(* IEC 61131-3 sources: plc-st-coding-agent/progress/evidence/f14_v11_public_20261113/jobs/custom_deepseek-v4pro (part 3) *)

(* ---- public-hard-04.raw_candidate_04.st ---- *)
(* ENGINEERING_CONTRACT
   elementCount DINT: retained process value; 0 after reset, +1 successful enqueue, -1 successful dequeue, held otherwise; range 0..capacity.
   status WORD: overwritten every invocation; 0 idle/reset/success, 16#8002 rejected full enqueue, 16#8001 rejected empty dequeue; reset priority sets 0.
   queue state: first invocation empty; reset priority clears head/tail/count; enqueue writes at tail, dequeue reads head; indices 0..capacity-1.
   edge triggers: R_TRIG consumed every scan; reset priority ignores edge requests; simultaneous enqueue+dequeue unspecified -> no-op.
   units/boundaries: capacity positive DINT derived once from buffer size / item element size; element copied byte-wise from item address.
*)
(* CONTRACT_RULES [] *)
FUNCTION_BLOCK FIFO
VAR_INPUT
    enqueue : BOOL;
    dequeue : BOOL;
    reset : BOOL;
END_VAR
VAR_OUTPUT
    elementCount : DINT;
    status : WORD;
END_VAR
VAR_IN_OUT
    item : VARIANT;
    buffer : VARIANT;
END_VAR
VAR
    local_rEnq : R_TRIG;
    local_rDeq : R_TRIG;
    local_enqEdge : BOOL;
    local_deqEdge : BOOL;

    local_associated : BOOL := FALSE;
    local_pBufferBase : POINTER TO BYTE;
    local_pItemBase : POINTER TO BYTE;
    local_elemSize : DINT := 1;
    local_capacity : DINT := 1;

    local_count : DINT := 0;
    local_head : DINT := 0;
    local_tail : DINT := 0;

    local_bufInfo : __SYSTEM.VAR_INFO;
    local_itemInfo : __SYSTEM.VAR_INFO;

    local_pSrc : POINTER TO BYTE;
    local_pDst : POINTER TO BYTE;
    local_offset : DINT;
    local_copiedBytes : UDINT;
END_VAR

(* Consume rising edges every scan so reset cannot create ghost operations later. *)
local_rEnq(CLK := enqueue);
local_enqEdge := local_rEnq.Q;
local_rDeq(CLK := dequeue);
local_deqEdge := local_rDeq.Q;

status := 16#0000;

(* One-time association of buffer and item storage, using the first invocation. *)
IF NOT local_associated THEN
    local_bufInfo := __VARINFO(buffer);
    local_itemInfo := __VARINFO(item);

    local_elemSize := local_itemInfo.diSize;
    IF local_elemSize <= 0 THEN
        local_elemSize := 1;
    END_IF;

    local_capacity := local_bufInfo.diSize / local_elemSize;
    IF local_capacity < 1 THEN
        local_capacity := 1;
    END_IF;

    local_pBufferBase := local_bufInfo.pvAddress;
    local_pItemBase := local_itemInfo.pvAddress;
    local_associated := TRUE;
END_IF;

IF reset THEN
    (* Reset has priority over all operations; stored values remain untouched. *)
    local_count := 0;
    local_head := 0;
    local_tail := 0;
    status := 16#0000;
ELSE
    IF local_enqEdge AND NOT local_deqEdge THEN
        IF local_count < local_capacity THEN
            (* Copy current item value into tail slot. *)
            local_pSrc := local_pItemBase;
            local_pDst := local_pBufferBase;
            local_offset := local_tail * local_elemSize;
            local_pDst := local_pDst + local_offset;
            local_copiedBytes := SysMemCpy(
                pbyDest := local_pDst,
                pbySource := local_pSrc,
                dwCount := TO_DWORD(local_elemSize)
            );

            local_tail := (local_tail + 1) MOD local_capacity;
            local_count := local_count + 1;
            status := 16#0000;
        ELSE
            status := 16#8002; (* enqueue rejected: full *)
        END_IF;
    ELSIF local_deqEdge AND NOT local_enqEdge THEN
        IF local_count > 0 THEN
            (* Copy head element back to item. *)
            local_pSrc := local_pBufferBase;
            local_offset := local_head * local_elemSize;
            local_pSrc := local_pSrc + local_offset;
            local_pDst := local_pItemBase;
            local_copiedBytes := SysMemCpy(
                pbyDest := local_pDst,
                pbySource := local_pSrc,
                dwCount := TO_DWORD(local_elemSize)
            );

            local_head := (local_head + 1) MOD local_capacity;
            local_count := local_count - 1;
            status := 16#0000;
        ELSE
            status := 16#8001; (* dequeue rejected: empty *)
        END_IF;
    END_IF;
END_IF;

elementCount := local_count;
END_FUNCTION_BLOCK

(* ---- public-hard-05.candidate_01.st ---- *)
(* ENGINEERING_CONTRACT
Manual: moving/grip/release outputs are combinational from corresponding button AND NOT corresponding limit switch; releasing the button clears the output. PUB001, PUB005.
SingleStep: rising Start advances only when idle or current step limit reached; each step holds its output until its limit, then waits for next Start. After step 8, next Start goes to step 1. PUB002.
SingleCycle: rising Start starts step 1; each step auto-advances on its completion limit, then stops at step 0 after step 8. PUB003.
Continuous: rising Start starts step 1; auto-advances and loops 8->1. PUB004.
EmergencyStop=FALSE forces all outputs FALSE and freezes automatic state changes. No reset is inferred. PUB005.
Completion feedback uses DownLimitSwitch, UpLimitSwitch, LeftLimitSwitch, RightLimitSwitch, GripLimitSwitch, ReleaseLimitSwitch. Unspecified mode-change behavior preserves the automatic step state.
*)
(* CONTRACT_RULES [] *)
FUNCTION_BLOCK FB_MechanicalArmControl
VAR CONSTANT
    cStepDown1 : INT := 1;
    cStepGrip : INT := 2;
    cStepUp1 : INT := 3;
    cStepRight : INT := 4;
    cStepDown2 : INT := 5;
    cStepRelease : INT := 6;
    cStepUp2 : INT := 7;
    cStepLeft : INT := 8;
END_VAR
VAR
    startTrig : R_TRIG;
    sdStep : INT := 0;
    autoStep : INT := 0;
    sdDone : BOOL;
    autoDone : BOOL;
    tmpMoveDown : BOOL;
    tmpMoveUp : BOOL;
    tmpMoveLeft : BOOL;
    tmpMoveRight : BOOL;
    tmpActivateGrip : BOOL;
    tmpActivateRelease : BOOL;
END_VAR

startTrig(CLK := Start);

tmpMoveDown := FALSE;
tmpMoveUp := FALSE;
tmpMoveLeft := FALSE;
tmpMoveRight := FALSE;
tmpActivateGrip := FALSE;
tmpActivateRelease := FALSE;

IF ManualMode THEN
    tmpMoveDown := DownButton AND NOT DownLimitSwitch;
    tmpMoveUp := UpButton AND NOT UpLimitSwitch;
    tmpMoveLeft := LeftButton AND NOT LeftLimitSwitch;
    tmpMoveRight := RightButton AND NOT RightLimitSwitch;
    tmpActivateGrip := GripButton AND NOT GripLimitSwitch;
    tmpActivateRelease := ReleaseButton AND NOT ReleaseLimitSwitch;

ELSIF SingleStepMode THEN
    CASE sdStep OF
        cStepDown1: sdDone := DownLimitSwitch;
        cStepGrip: sdDone := GripLimitSwitch;
        cStepUp1: sdDone := UpLimitSwitch;
        cStepRight: sdDone := RightLimitSwitch;
        cStepDown2: sdDone := DownLimitSwitch;
        cStepRelease: sdDone := ReleaseLimitSwitch;
        cStepUp2: sdDone := UpLimitSwitch;
        cStepLeft: sdDone := LeftLimitSwitch;
    ELSE
        sdDone := TRUE;
    END_CASE;

    IF EmergencyStop AND startTrig.Q AND sdDone THEN
        IF sdStep >= cStepLeft THEN
            sdStep := cStepDown1;
        ELSE
            sdStep := sdStep + 1;
        END_IF;
    END_IF;

    CASE sdStep OF
        cStepDown1: tmpMoveDown := NOT DownLimitSwitch;
        cStepGrip: tmpActivateGrip := NOT GripLimitSwitch;
        cStepUp1: tmpMoveUp := NOT UpLimitSwitch;
        cStepRight: tmpMoveRight := NOT RightLimitSwitch;
        cStepDown2: tmpMoveDown := NOT DownLimitSwitch;
        cStepRelease: tmpActivateRelease := NOT ReleaseLimitSwitch;
        cStepUp2: tmpMoveUp := NOT UpLimitSwitch;
        cStepLeft: tmpMoveLeft := NOT LeftLimitSwitch;
    ELSE
        // no automatic output
    END_CASE;

ELSIF SingleCycleMode OR ContinuousMode THEN
    IF EmergencyStop AND startTrig.Q AND (autoStep = 0) THEN
        autoStep := cStepDown1;
    END_IF;

    CASE autoStep OF
        cStepDown1: autoDone := DownLimitSwitch;
        cStepGrip: autoDone := GripLimitSwitch;
        cStepUp1: autoDone := UpLimitSwitch;
        cStepRight: autoDone := RightLimitSwitch;
        cStepDown2: autoDone := DownLimitSwitch;
        cStepRelease: autoDone := ReleaseLimitSwitch;
        cStepUp2: autoDone := UpLimitSwitch;
        cStepLeft: autoDone := LeftLimitSwitch;
    ELSE
        autoDone := TRUE;
    END_CASE;

    IF EmergencyStop AND (autoStep <> 0) AND autoDone THEN
        IF SingleCycleMode THEN
            IF autoStep < cStepLeft THEN
                autoStep := autoStep + 1;
            ELSE
                autoStep := 0;
            END_IF;
        ELSIF ContinuousMode THEN
            IF autoStep < cStepLeft THEN
                autoStep := autoStep + 1;
            ELSE
                autoStep := cStepDown1;
            END_IF;
        END_IF;
    END_IF;

    CASE autoStep OF
        cStepDown1: tmpMoveDown := NOT DownLimitSwitch;
        cStepGrip: tmpActivateGrip := NOT GripLimitSwitch;
        cStepUp1: tmpMoveUp := NOT UpLimitSwitch;
        cStepRight: tmpMoveRight := NOT RightLimitSwitch;
        cStepDown2: tmpMoveDown := NOT DownLimitSwitch;
        cStepRelease: tmpActivateRelease := NOT ReleaseLimitSwitch;
        cStepUp2: tmpMoveUp := NOT UpLimitSwitch;
        cStepLeft: tmpMoveLeft := NOT LeftLimitSwitch;
    ELSE
        // idle/no output
    END_CASE;
END_IF;

IF NOT EmergencyStop THEN
    MoveDown := FALSE;
    MoveUp := FALSE;
    MoveLeft := FALSE;
    MoveRight := FALSE;
    ActivateGrip := FALSE;
    ActivateRelease := FALSE;
ELSE
    MoveDown := tmpMoveDown;
    MoveUp := tmpMoveUp;
    MoveLeft := tmpMoveLeft;
    MoveRight := tmpMoveRight;
    ActivateGrip := tmpActivateGrip;
    ActivateRelease := tmpActivateRelease;
END_IF;

END_FUNCTION_BLOCK

(* ---- public-hard-05.candidate_02.st ---- *)
(* ENGINEERING_CONTRACT
Manual: moving/grip/release outputs are combinational from corresponding button AND NOT corresponding limit switch; releasing the button clears the output. PUB001, PUB005.
SingleStep: rising Start advances only when idle or current step limit reached; each step holds its output until its limit, then waits for next Start. After step 8, next Start goes to step 1. PUB002.
SingleCycle: rising Start starts step 1; each step auto-advances on its completion limit, then stops at step 0 after step 8. PUB003.
Continuous: rising Start starts step 1; auto-advances and loops 8->1. PUB004.
EmergencyStop=FALSE forces all outputs FALSE and freezes automatic state changes. No reset is inferred. PUB005.
Completion feedback uses DownLimitSwitch, UpLimitSwitch, LeftLimitSwitch, RightLimitSwitch, GripLimitSwitch, ReleaseLimitSwitch. Unspecified mode-change behavior preserves the automatic step state.
*)
(* CONTRACT_RULES [] *)
FUNCTION_BLOCK FB_MechanicalArmControl
VAR CONSTANT
    cStepDown1 : INT := 1;
    cStepGrip : INT := 2;
    cStepUp1 : INT := 3;
    cStepRight : INT := 4;
    cStepDown2 : INT := 5;
    cStepRelease : INT := 6;
    cStepUp2 : INT := 7;
    cStepLeft : INT := 8;
END_VAR
VAR
    startTrig : R_TRIG;
    sdStep : INT := 0;
    autoStep : INT := 0;
    sdDone : BOOL;
    autoDone : BOOL;
    tmpMoveDown : BOOL;
    tmpMoveUp : BOOL;
    tmpMoveLeft : BOOL;
    tmpMoveRight : BOOL;
    tmpActivateGrip : BOOL;
    tmpActivateRelease : BOOL;
END_VAR

startTrig(CLK := Start);

tmpMoveDown := FALSE;
tmpMoveUp := FALSE;
tmpMoveLeft := FALSE;
tmpMoveRight := FALSE;
tmpActivateGrip := FALSE;
tmpActivateRelease := FALSE;

IF ManualMode THEN
    tmpMoveDown := DownButton AND NOT DownLimitSwitch;
    tmpMoveUp := UpButton AND NOT UpLimitSwitch;
    tmpMoveLeft := LeftButton AND NOT LeftLimitSwitch;
    tmpMoveRight := RightButton AND NOT RightLimitSwitch;
    tmpActivateGrip := GripButton AND NOT GripLimitSwitch;
    tmpActivateRelease := ReleaseButton AND NOT ReleaseLimitSwitch;

ELSIF SingleStepMode THEN
    CASE sdStep OF
        cStepDown1: sdDone := DownLimitSwitch;
        cStepGrip: sdDone := GripLimitSwitch;
        cStepUp1: sdDone := UpLimitSwitch;
        cStepRight: sdDone := RightLimitSwitch;
        cStepDown2: sdDone := DownLimitSwitch;
        cStepRelease: sdDone := ReleaseLimitSwitch;
        cStepUp2: sdDone := UpLimitSwitch;
        cStepLeft: sdDone := LeftLimitSwitch;
    ELSE
        sdDone := TRUE;
    END_CASE;

    IF EmergencyStop AND startTrig.Q AND sdDone THEN
        IF sdStep >= cStepLeft THEN
            sdStep := cStepDown1;
        ELSE
            sdStep := sdStep + 1;
        END_IF;
    END_IF;

    CASE sdStep OF
        cStepDown1: tmpMoveDown := NOT DownLimitSwitch;
        cStepGrip: tmpActivateGrip := NOT GripLimitSwitch;
        cStepUp1: tmpMoveUp := NOT UpLimitSwitch;
        cStepRight: tmpMoveRight := NOT RightLimitSwitch;
        cStepDown2: tmpMoveDown := NOT DownLimitSwitch;
        cStepRelease: tmpActivateRelease := NOT ReleaseLimitSwitch;
        cStepUp2: tmpMoveUp := NOT UpLimitSwitch;
        cStepLeft: tmpMoveLeft := NOT LeftLimitSwitch;
    ELSE
        (* no automatic output *)
    END_CASE;

ELSIF SingleCycleMode OR ContinuousMode THEN
    IF EmergencyStop AND startTrig.Q AND (autoStep = 0) THEN
        autoStep := cStepDown1;
    END_IF;

    CASE autoStep OF
        cStepDown1: autoDone := DownLimitSwitch;
        cStepGrip: autoDone := GripLimitSwitch;
        cStepUp1: autoDone := UpLimitSwitch;
        cStepRight: autoDone := RightLimitSwitch;
        cStepDown2: autoDone := DownLimitSwitch;
        cStepRelease: autoDone := ReleaseLimitSwitch;
        cStepUp2: autoDone := UpLimitSwitch;
        cStepLeft: autoDone := LeftLimitSwitch;
    ELSE
        autoDone := TRUE;
    END_CASE;

    IF EmergencyStop AND (autoStep <> 0) AND autoDone THEN
        IF SingleCycleMode THEN
            IF autoStep < cStepLeft THEN
                autoStep := autoStep + 1;
            ELSE
                autoStep := 0;
            END_IF;
        ELSIF ContinuousMode THEN
            IF autoStep < cStepLeft THEN
                autoStep := autoStep + 1;
            ELSE
                autoStep := cStepDown1;
            END_IF;
        END_IF;
    END_IF;

    CASE autoStep OF
        cStepDown1: tmpMoveDown := NOT DownLimitSwitch;
        cStepGrip: tmpActivateGrip := NOT GripLimitSwitch;
        cStepUp1: tmpMoveUp := NOT UpLimitSwitch;
        cStepRight: tmpMoveRight := NOT RightLimitSwitch;
        cStepDown2: tmpMoveDown := NOT DownLimitSwitch;
        cStepRelease: tmpActivateRelease := NOT ReleaseLimitSwitch;
        cStepUp2: tmpMoveUp := NOT UpLimitSwitch;
        cStepLeft: tmpMoveLeft := NOT LeftLimitSwitch;
    ELSE
        (* idle/no output *)
    END_CASE;
END_IF;

IF NOT EmergencyStop THEN
    MoveDown := FALSE;
    MoveUp := FALSE;
    MoveLeft := FALSE;
    MoveRight := FALSE;
    ActivateGrip := FALSE;
    ActivateRelease := FALSE;
ELSE
    MoveDown := tmpMoveDown;
    MoveUp := tmpMoveUp;
    MoveLeft := tmpMoveLeft;
    MoveRight := tmpMoveRight;
    ActivateGrip := tmpActivateGrip;
    ActivateRelease := tmpActivateRelease;
END_IF;

END_FUNCTION_BLOCK

(* ---- public-hard-05.candidate_03.st ---- *)
(* ENGINEERING_CONTRACT
Manual: moving/grip/release outputs are combinational from corresponding button AND NOT corresponding limit switch; releasing the button clears the output. PUB001, PUB005.
SingleStep: rising Start advances only when idle or current step limit reached; each step holds its output until its limit, then waits for next Start. After step 8, next Start goes to step 1. PUB002.
SingleCycle: rising Start starts step 1; each step auto-advances on its completion limit, then stops at step 0 after step 8. PUB003.
Continuous: rising Start starts step 1; auto-advances and loops 8->1. PUB004.
EmergencyStop=FALSE forces all outputs FALSE and freezes automatic state changes. No reset is inferred. PUB005.
Completion feedback uses DownLimitSwitch, UpLimitSwitch, LeftLimitSwitch, RightLimitSwitch, GripLimitSwitch, ReleaseLimitSwitch. Unspecified mode-change behavior preserves the automatic step state.
*)
(* CONTRACT_RULES [] *)
FUNCTION_BLOCK FB_MechanicalArmControl
VAR CONSTANT
    cStepDown1 : INT := 1;
    cStepGrip : INT := 2;
    cStepUp1 : INT := 3;
    cStepRight : INT := 4;
    cStepDown2 : INT := 5;
    cStepRelease : INT := 6;
    cStepUp2 : INT := 7;
    cStepLeft : INT := 8;
END_VAR
VAR_INPUT
    ManualMode : BOOL;
    SingleStepMode : BOOL;
    SingleCycleMode : BOOL;
    ContinuousMode : BOOL;
    EmergencyStop : BOOL;
    Start : BOOL;
    DownButton : BOOL;
    UpButton : BOOL;
    LeftButton : BOOL;
    RightButton : BOOL;
    GripButton : BOOL;
    ReleaseButton : BOOL;
    DownLimitSwitch : BOOL;
    UpLimitSwitch : BOOL;
    LeftLimitSwitch : BOOL;
    RightLimitSwitch : BOOL;
    GripLimitSwitch : BOOL;
    ReleaseLimitSwitch : BOOL;
END_VAR
VAR_OUTPUT
    MoveDown : BOOL;
    MoveUp : BOOL;
    MoveLeft : BOOL;
    MoveRight : BOOL;
    ActivateGrip : BOOL;
    ActivateRelease : BOOL;
END_VAR
VAR
    startTrig : R_TRIG;
    sdStep : INT := 0;
    autoStep : INT := 0;
    sdDone : BOOL;
    autoDone : BOOL;
    tmpMoveDown : BOOL;
    tmpMoveUp : BOOL;
    tmpMoveLeft : BOOL;
    tmpMoveRight : BOOL;
    tmpActivateGrip : BOOL;
    tmpActivateRelease : BOOL;
END_VAR

startTrig(CLK := Start);

tmpMoveDown := FALSE;
tmpMoveUp := FALSE;
tmpMoveLeft := FALSE;
tmpMoveRight := FALSE;
tmpActivateGrip := FALSE;
tmpActivateRelease := FALSE;

IF ManualMode THEN
    tmpMoveDown := DownButton AND NOT DownLimitSwitch;
    tmpMoveUp := UpButton AND NOT UpLimitSwitch;
    tmpMoveLeft := LeftButton AND NOT LeftLimitSwitch;
    tmpMoveRight := RightButton AND NOT RightLimitSwitch;
    tmpActivateGrip := GripButton AND NOT GripLimitSwitch;
    tmpActivateRelease := ReleaseButton AND NOT ReleaseLimitSwitch;

ELSIF SingleStepMode THEN
    CASE sdStep OF
        cStepDown1: sdDone := DownLimitSwitch;
        cStepGrip: sdDone := GripLimitSwitch;
        cStepUp1: sdDone := UpLimitSwitch;
        cStepRight: sdDone := RightLimitSwitch;
        cStepDown2: sdDone := DownLimitSwitch;
        cStepRelease: sdDone := ReleaseLimitSwitch;
        cStepUp2: sdDone := UpLimitSwitch;
        cStepLeft: sdDone := LeftLimitSwitch;
    ELSE
        sdDone := TRUE;
    END_CASE;

    IF EmergencyStop AND startTrig.Q AND sdDone THEN
        IF sdStep >= cStepLeft THEN
            sdStep := cStepDown1;
        ELSE
            sdStep := sdStep + 1;
        END_IF;
    END_IF;

    CASE sdStep OF
        cStepDown1: tmpMoveDown := NOT DownLimitSwitch;
        cStepGrip: tmpActivateGrip := NOT GripLimitSwitch;
        cStepUp1: tmpMoveUp := NOT UpLimitSwitch;
        cStepRight: tmpMoveRight := NOT RightLimitSwitch;
        cStepDown2: tmpMoveDown := NOT DownLimitSwitch;
        cStepRelease: tmpActivateRelease := NOT ReleaseLimitSwitch;
        cStepUp2: tmpMoveUp := NOT UpLimitSwitch;
        cStepLeft: tmpMoveLeft := NOT LeftLimitSwitch;
    ELSE
        (* no automatic output *)
    END_CASE;

ELSIF SingleCycleMode OR ContinuousMode THEN
    IF EmergencyStop AND startTrig.Q AND (autoStep = 0) THEN
        autoStep := cStepDown1;
    END_IF;

    CASE autoStep OF
        cStepDown1: autoDone := DownLimitSwitch;
        cStepGrip: autoDone := GripLimitSwitch;
        cStepUp1: autoDone := UpLimitSwitch;
        cStepRight: autoDone := RightLimitSwitch;
        cStepDown2: autoDone := DownLimitSwitch;
        cStepRelease: autoDone := ReleaseLimitSwitch;
        cStepUp2: autoDone := UpLimitSwitch;
        cStepLeft: autoDone := LeftLimitSwitch;
    ELSE
        autoDone := TRUE;
    END_CASE;

    IF EmergencyStop AND (autoStep <> 0) AND autoDone THEN
        IF SingleCycleMode THEN
            IF autoStep < cStepLeft THEN
                autoStep := autoStep + 1;
            ELSE
                autoStep := 0;
            END_IF;
        ELSIF ContinuousMode THEN
            IF autoStep < cStepLeft THEN
                autoStep := autoStep + 1;
            ELSE
                autoStep := cStepDown1;
            END_IF;
        END_IF;
    END_IF;

    CASE autoStep OF
        cStepDown1: tmpMoveDown := NOT DownLimitSwitch;
        cStepGrip: tmpActivateGrip := NOT GripLimitSwitch;
        cStepUp1: tmpMoveUp := NOT UpLimitSwitch;
        cStepRight: tmpMoveRight := NOT RightLimitSwitch;
        cStepDown2: tmpMoveDown := NOT DownLimitSwitch;
        cStepRelease: tmpActivateRelease := NOT ReleaseLimitSwitch;
        cStepUp2: tmpMoveUp := NOT UpLimitSwitch;
        cStepLeft: tmpMoveLeft := NOT LeftLimitSwitch;
    ELSE
        (* idle/no output *)
    END_CASE;

END_IF;

IF NOT EmergencyStop THEN
    MoveDown := FALSE;
    MoveUp := FALSE;
    MoveLeft := FALSE;
    MoveRight := FALSE;
    ActivateGrip := FALSE;
    ActivateRelease := FALSE;
ELSE
    MoveDown := tmpMoveDown;
    MoveUp := tmpMoveUp;
    MoveLeft := tmpMoveLeft;
    MoveRight := tmpMoveRight;
    ActivateGrip := tmpActivateGrip;
    ActivateRelease := tmpActivateRelease;
END_IF;

END_FUNCTION_BLOCK

(* ---- public-hard-05.candidate_04.st ---- *)
(* ENGINEERING_CONTRACT
Manual: moving/grip/release outputs are combinational from corresponding button AND NOT corresponding limit switch; releasing the button clears the output. PUB001, PUB005.
SingleStep: rising Start advances only when idle or current step limit reached; each step holds its output until its limit, then waits for next Start. After step 8, next Start goes to step 1. PUB002.
SingleCycle: rising Start starts step 1; each step auto-advances on its completion limit, then stops at step 0 after step 8. PUB003.
Continuous: rising Start starts step 1; auto-advances and loops 8->1. PUB004.
EmergencyStop=FALSE forces all outputs FALSE and freezes automatic state changes. No reset is inferred. PUB005.
Completion feedback uses DownLimitSwitch, UpLimitSwitch, LeftLimitSwitch, RightLimitSwitch, GripLimitSwitch, ReleaseLimitSwitch. Unspecified mode-change behavior preserves the automatic step state.
*)
(* CONTRACT_RULES [] *)
FUNCTION_BLOCK FB_MechanicalArmControl
VAR_INPUT
    ManualMode : BOOL;
    SingleStepMode : BOOL;
    SingleCycleMode : BOOL;
    ContinuousMode : BOOL;
    EmergencyStop : BOOL;
    Start : BOOL;
    DownButton : BOOL;
    UpButton : BOOL;
    LeftButton : BOOL;
    RightButton : BOOL;
    GripButton : BOOL;
    ReleaseButton : BOOL;
    DownLimitSwitch : BOOL;
    UpLimitSwitch : BOOL;
    LeftLimitSwitch : BOOL;
    RightLimitSwitch : BOOL;
    GripLimitSwitch : BOOL;
    ReleaseLimitSwitch : BOOL;
END_VAR
VAR_OUTPUT
    MoveDown : BOOL;
    MoveUp : BOOL;
    MoveLeft : BOOL;
    MoveRight : BOOL;
    ActivateGrip : BOOL;
    ActivateRelease : BOOL;
END_VAR
VAR
    startTrig : R_TRIG;
    sdStep : INT := 0;
    autoStep : INT := 0;
    sdDone : BOOL;
    autoDone : BOOL;
    tmpMoveDown : BOOL;
    tmpMoveUp : BOOL;
    tmpMoveLeft : BOOL;
    tmpMoveRight : BOOL;
    tmpActivateGrip : BOOL;
    tmpActivateRelease : BOOL;
END_VAR

startTrig(CLK := Start);

tmpMoveDown := FALSE;
tmpMoveUp := FALSE;
tmpMoveLeft := FALSE;
tmpMoveRight := FALSE;
tmpActivateGrip := FALSE;
tmpActivateRelease := FALSE;

IF ManualMode THEN
    tmpMoveDown := DownButton AND NOT DownLimitSwitch;
    tmpMoveUp := UpButton AND NOT UpLimitSwitch;
    tmpMoveLeft := LeftButton AND NOT LeftLimitSwitch;
    tmpMoveRight := RightButton AND NOT RightLimitSwitch;
    tmpActivateGrip := GripButton AND NOT GripLimitSwitch;
    tmpActivateRelease := ReleaseButton AND NOT ReleaseLimitSwitch;

ELSIF SingleStepMode THEN
    CASE sdStep OF
        1: sdDone := DownLimitSwitch;
        2: sdDone := GripLimitSwitch;
        3: sdDone := UpLimitSwitch;
        4: sdDone := RightLimitSwitch;
        5: sdDone := DownLimitSwitch;
        6: sdDone := ReleaseLimitSwitch;
        7: sdDone := UpLimitSwitch;
        8: sdDone := LeftLimitSwitch;
    ELSE
        sdDone := TRUE;
    END_CASE;

    IF EmergencyStop AND startTrig.Q AND sdDone THEN
        IF sdStep >= 8 THEN
            sdStep := 1;
        ELSE
            sdStep := sdStep + 1;
        END_IF;
    END_IF;

    CASE sdStep OF
        1: tmpMoveDown := NOT DownLimitSwitch;
        2: tmpActivateGrip := NOT GripLimitSwitch;
        3: tmpMoveUp := NOT UpLimitSwitch;
        4: tmpMoveRight := NOT RightLimitSwitch;
        5: tmpMoveDown := NOT DownLimitSwitch;
        6: tmpActivateRelease := NOT ReleaseLimitSwitch;
        7: tmpMoveUp := NOT UpLimitSwitch;
        8: tmpMoveLeft := NOT LeftLimitSwitch;
    END_CASE;

ELSIF (SingleCycleMode OR ContinuousMode) THEN
    IF EmergencyStop AND startTrig.Q AND (autoStep = 0) THEN
        autoStep := 1;
    END_IF;

    CASE autoStep OF
        1: autoDone := DownLimitSwitch;
        2: autoDone := GripLimitSwitch;
        3: autoDone := UpLimitSwitch;
        4: autoDone := RightLimitSwitch;
        5: autoDone := DownLimitSwitch;
        6: autoDone := ReleaseLimitSwitch;
        7: autoDone := UpLimitSwitch;
        8: autoDone := LeftLimitSwitch;
    ELSE
        autoDone := TRUE;
    END_CASE;

    IF EmergencyStop AND (autoStep <> 0) AND autoDone THEN
        IF SingleCycleMode THEN
            IF autoStep < 8 THEN
                autoStep := autoStep + 1;
            ELSE
                autoStep := 0;
            END_IF;
        ELSIF ContinuousMode THEN
            IF autoStep < 8 THEN
                autoStep := autoStep + 1;
            ELSE
                autoStep := 1;
            END_IF;
        END_IF;
    END_IF;

    CASE autoStep OF
        1: tmpMoveDown := NOT DownLimitSwitch;
        2: tmpActivateGrip := NOT GripLimitSwitch;
        3: tmpMoveUp := NOT UpLimitSwitch;
        4: tmpMoveRight := NOT RightLimitSwitch;
        5: tmpMoveDown := NOT DownLimitSwitch;
        6: tmpActivateRelease := NOT ReleaseLimitSwitch;
        7: tmpMoveUp := NOT UpLimitSwitch;
        8: tmpMoveLeft := NOT LeftLimitSwitch;
    END_CASE;

END_IF;

IF NOT EmergencyStop THEN
    MoveDown := FALSE;
    MoveUp := FALSE;
    MoveLeft := FALSE;
    MoveRight := FALSE;
    ActivateGrip := FALSE;
    ActivateRelease := FALSE;
ELSE
    MoveDown := tmpMoveDown;
    MoveUp := tmpMoveUp;
    MoveLeft := tmpMoveLeft;
    MoveRight := tmpMoveRight;
    ActivateGrip := tmpActivateGrip;
    ActivateRelease := tmpActivateRelease;
END_IF;

END_FUNCTION_BLOCK

(* ---- public-hard-05.raw_candidate_01.st ---- *)
(* ENGINEERING_CONTRACT
Manual: moving/grip/release outputs are combinational from corresponding button AND NOT corresponding limit switch; releasing the button clears the output. PUB001, PUB005.
SingleStep: rising Start advances only when idle or current step limit reached; each step holds its output until its limit, then waits for next Start. After step 8, next Start goes to step 1. PUB002.
SingleCycle: rising Start starts step 1; each step auto-advances on its completion limit, then stops at step 0 after step 8. PUB003.
Continuous: rising Start starts step 1; auto-advances and loops 8->1. PUB004.
EmergencyStop=FALSE forces all outputs FALSE and freezes automatic state changes. No reset is inferred. PUB005.
Completion feedback uses DownLimitSwitch, UpLimitSwitch, LeftLimitSwitch, RightLimitSwitch, GripLimitSwitch, ReleaseLimitSwitch. Unspecified mode-change behavior preserves the automatic step state.
*)
(* CONTRACT_RULES [] *)
FUNCTION_BLOCK FB_MechanicalArmControl
VAR CONSTANT
    cStepDown1 : INT := 1;
    cStepGrip : INT := 2;
    cStepUp1 : INT := 3;
    cStepRight : INT := 4;
    cStepDown2 : INT := 5;
    cStepRelease : INT := 6;
    cStepUp2 : INT := 7;
    cStepLeft : INT := 8;
END_VAR
VAR
    startTrig : R_TRIG;
    sdStep : INT := 0;
    autoStep : INT := 0;
    sdDone : BOOL;
    autoDone : BOOL;
    tmpMoveDown : BOOL;
    tmpMoveUp : BOOL;
    tmpMoveLeft : BOOL;
    tmpMoveRight : BOOL;
    tmpActivateGrip : BOOL;
    tmpActivateRelease : BOOL;
END_VAR

startTrig(CLK := Start);

tmpMoveDown := FALSE;
tmpMoveUp := FALSE;
tmpMoveLeft := FALSE;
tmpMoveRight := FALSE;
tmpActivateGrip := FALSE;
tmpActivateRelease := FALSE;

IF ManualMode THEN
    tmpMoveDown := DownButton AND NOT DownLimitSwitch;
    tmpMoveUp := UpButton AND NOT UpLimitSwitch;
    tmpMoveLeft := LeftButton AND NOT LeftLimitSwitch;
    tmpMoveRight := RightButton AND NOT RightLimitSwitch;
    tmpActivateGrip := GripButton AND NOT GripLimitSwitch;
    tmpActivateRelease := ReleaseButton AND NOT ReleaseLimitSwitch;

ELSIF SingleStepMode THEN
    CASE sdStep OF
        cStepDown1: sdDone := DownLimitSwitch;
        cStepGrip: sdDone := GripLimitSwitch;
        cStepUp1: sdDone := UpLimitSwitch;
        cStepRight: sdDone := RightLimitSwitch;
        cStepDown2: sdDone := DownLimitSwitch;
        cStepRelease: sdDone := ReleaseLimitSwitch;
        cStepUp2: sdDone := UpLimitSwitch;
        cStepLeft: sdDone := LeftLimitSwitch;
    ELSE
        sdDone := TRUE;
    END_CASE;

    IF EmergencyStop AND startTrig.Q AND sdDone THEN
        IF sdStep >= cStepLeft THEN
            sdStep := cStepDown1;
        ELSE
            sdStep := sdStep + 1;
        END_IF;
    END_IF;

    CASE sdStep OF
        cStepDown1: tmpMoveDown := NOT DownLimitSwitch;
        cStepGrip: tmpActivateGrip := NOT GripLimitSwitch;
        cStepUp1: tmpMoveUp := NOT UpLimitSwitch;
        cStepRight: tmpMoveRight := NOT RightLimitSwitch;
        cStepDown2: tmpMoveDown := NOT DownLimitSwitch;
        cStepRelease: tmpActivateRelease := NOT ReleaseLimitSwitch;
        cStepUp2: tmpMoveUp := NOT UpLimitSwitch;
        cStepLeft: tmpMoveLeft := NOT LeftLimitSwitch;
    ELSE
        // no automatic output
    END_CASE;

ELSIF SingleCycleMode OR ContinuousMode THEN
    IF EmergencyStop AND startTrig.Q AND (autoStep = 0) THEN
        autoStep := cStepDown1;
    END_IF;

    CASE autoStep OF
        cStepDown1: autoDone := DownLimitSwitch;
        cStepGrip: autoDone := GripLimitSwitch;
        cStepUp1: autoDone := UpLimitSwitch;
        cStepRight: autoDone := RightLimitSwitch;
        cStepDown2: autoDone := DownLimitSwitch;
        cStepRelease: autoDone := ReleaseLimitSwitch;
        cStepUp2: autoDone := UpLimitSwitch;
        cStepLeft: autoDone := LeftLimitSwitch;
    ELSE
        autoDone := TRUE;
    END_CASE;

    IF EmergencyStop AND (autoStep <> 0) AND autoDone THEN
        IF SingleCycleMode THEN
            IF autoStep < cStepLeft THEN
                autoStep := autoStep + 1;
            ELSE
                autoStep := 0;
            END_IF;
        ELSIF ContinuousMode THEN
            IF autoStep < cStepLeft THEN
                autoStep := autoStep + 1;
            ELSE
                autoStep := cStepDown1;
            END_IF;
        END_IF;
    END_IF;

    CASE autoStep OF
        cStepDown1: tmpMoveDown := NOT DownLimitSwitch;
        cStepGrip: tmpActivateGrip := NOT GripLimitSwitch;
        cStepUp1: tmpMoveUp := NOT UpLimitSwitch;
        cStepRight: tmpMoveRight := NOT RightLimitSwitch;
        cStepDown2: tmpMoveDown := NOT DownLimitSwitch;
        cStepRelease: tmpActivateRelease := NOT ReleaseLimitSwitch;
        cStepUp2: tmpMoveUp := NOT UpLimitSwitch;
        cStepLeft: tmpMoveLeft := NOT LeftLimitSwitch;
    ELSE
        // idle/no output
    END_CASE;
END_IF;

IF NOT EmergencyStop THEN
    MoveDown := FALSE;
    MoveUp := FALSE;
    MoveLeft := FALSE;
    MoveRight := FALSE;
    ActivateGrip := FALSE;
    ActivateRelease := FALSE;
ELSE
    MoveDown := tmpMoveDown;
    MoveUp := tmpMoveUp;
    MoveLeft := tmpMoveLeft;
    MoveRight := tmpMoveRight;
    ActivateGrip := tmpActivateGrip;
    ActivateRelease := tmpActivateRelease;
END_IF;

END_FUNCTION_BLOCK

(* ---- public-hard-05.raw_candidate_02.st ---- *)
(* ENGINEERING_CONTRACT
Manual: moving/grip/release outputs are combinational from corresponding button AND NOT corresponding limit switch; releasing the button clears the output. PUB001, PUB005.
SingleStep: rising Start advances only when idle or current step limit reached; each step holds its output until its limit, then waits for next Start. After step 8, next Start goes to step 1. PUB002.
SingleCycle: rising Start starts step 1; each step auto-advances on its completion limit, then stops at step 0 after step 8. PUB003.
Continuous: rising Start starts step 1; auto-advances and loops 8->1. PUB004.
EmergencyStop=FALSE forces all outputs FALSE and freezes automatic state changes. No reset is inferred. PUB005.
Completion feedback uses DownLimitSwitch, UpLimitSwitch, LeftLimitSwitch, RightLimitSwitch, GripLimitSwitch, ReleaseLimitSwitch. Unspecified mode-change behavior preserves the automatic step state.
*)
(* CONTRACT_RULES [] *)
FUNCTION_BLOCK FB_MechanicalArmControl
VAR CONSTANT
    cStepDown1 : INT := 1;
    cStepGrip : INT := 2;
    cStepUp1 : INT := 3;
    cStepRight : INT := 4;
    cStepDown2 : INT := 5;
    cStepRelease : INT := 6;
    cStepUp2 : INT := 7;
    cStepLeft : INT := 8;
END_VAR
VAR
    startTrig : R_TRIG;
    sdStep : INT := 0;
    autoStep : INT := 0;
    sdDone : BOOL;
    autoDone : BOOL;
    tmpMoveDown : BOOL;
    tmpMoveUp : BOOL;
    tmpMoveLeft : BOOL;
    tmpMoveRight : BOOL;
    tmpActivateGrip : BOOL;
    tmpActivateRelease : BOOL;
END_VAR

startTrig(CLK := Start);

tmpMoveDown := FALSE;
tmpMoveUp := FALSE;
tmpMoveLeft := FALSE;
tmpMoveRight := FALSE;
tmpActivateGrip := FALSE;
tmpActivateRelease := FALSE;

IF ManualMode THEN
    tmpMoveDown := DownButton AND NOT DownLimitSwitch;
    tmpMoveUp := UpButton AND NOT UpLimitSwitch;
    tmpMoveLeft := LeftButton AND NOT LeftLimitSwitch;
    tmpMoveRight := RightButton AND NOT RightLimitSwitch;
    tmpActivateGrip := GripButton AND NOT GripLimitSwitch;
    tmpActivateRelease := ReleaseButton AND NOT ReleaseLimitSwitch;

ELSIF SingleStepMode THEN
    CASE sdStep OF
        cStepDown1: sdDone := DownLimitSwitch;
        cStepGrip: sdDone := GripLimitSwitch;
        cStepUp1: sdDone := UpLimitSwitch;
        cStepRight: sdDone := RightLimitSwitch;
        cStepDown2: sdDone := DownLimitSwitch;
        cStepRelease: sdDone := ReleaseLimitSwitch;
        cStepUp2: sdDone := UpLimitSwitch;
        cStepLeft: sdDone := LeftLimitSwitch;
    ELSE
        sdDone := TRUE;
    END_CASE;

    IF EmergencyStop AND startTrig.Q AND sdDone THEN
        IF sdStep >= cStepLeft THEN
            sdStep := cStepDown1;
        ELSE
            sdStep := sdStep + 1;
        END_IF;
    END_IF;

    CASE sdStep OF
        cStepDown1: tmpMoveDown := NOT DownLimitSwitch;
        cStepGrip: tmpActivateGrip := NOT GripLimitSwitch;
        cStepUp1: tmpMoveUp := NOT UpLimitSwitch;
        cStepRight: tmpMoveRight := NOT RightLimitSwitch;
        cStepDown2: tmpMoveDown := NOT DownLimitSwitch;
        cStepRelease: tmpActivateRelease := NOT ReleaseLimitSwitch;
        cStepUp2: tmpMoveUp := NOT UpLimitSwitch;
        cStepLeft: tmpMoveLeft := NOT LeftLimitSwitch;
    ELSE
        (* no automatic output *)
    END_CASE;

ELSIF SingleCycleMode OR ContinuousMode THEN
    IF EmergencyStop AND startTrig.Q AND (autoStep = 0) THEN
        autoStep := cStepDown1;
    END_IF;

    CASE autoStep OF
        cStepDown1: autoDone := DownLimitSwitch;
        cStepGrip: autoDone := GripLimitSwitch;
        cStepUp1: autoDone := UpLimitSwitch;
        cStepRight: autoDone := RightLimitSwitch;
        cStepDown2: autoDone := DownLimitSwitch;
        cStepRelease: autoDone := ReleaseLimitSwitch;
        cStepUp2: autoDone := UpLimitSwitch;
        cStepLeft: autoDone := LeftLimitSwitch;
    ELSE
        autoDone := TRUE;
    END_CASE;

    IF EmergencyStop AND (autoStep <> 0) AND autoDone THEN
        IF SingleCycleMode THEN
            IF autoStep < cStepLeft THEN
                autoStep := autoStep + 1;
            ELSE
                autoStep := 0;
            END_IF;
        ELSIF ContinuousMode THEN
            IF autoStep < cStepLeft THEN
                autoStep := autoStep + 1;
            ELSE
                autoStep := cStepDown1;
            END_IF;
        END_IF;
    END_IF;

    CASE autoStep OF
        cStepDown1: tmpMoveDown := NOT DownLimitSwitch;
        cStepGrip: tmpActivateGrip := NOT GripLimitSwitch;
        cStepUp1: tmpMoveUp := NOT UpLimitSwitch;
        cStepRight: tmpMoveRight := NOT RightLimitSwitch;
        cStepDown2: tmpMoveDown := NOT DownLimitSwitch;
        cStepRelease: tmpActivateRelease := NOT ReleaseLimitSwitch;
        cStepUp2: tmpMoveUp := NOT UpLimitSwitch;
        cStepLeft: tmpMoveLeft := NOT LeftLimitSwitch;
    ELSE
        (* idle/no output *)
    END_CASE;
END_IF;

IF NOT EmergencyStop THEN
    MoveDown := FALSE;
    MoveUp := FALSE;
    MoveLeft := FALSE;
    MoveRight := FALSE;
    ActivateGrip := FALSE;
    ActivateRelease := FALSE;
ELSE
    MoveDown := tmpMoveDown;
    MoveUp := tmpMoveUp;
    MoveLeft := tmpMoveLeft;
    MoveRight := tmpMoveRight;
    ActivateGrip := tmpActivateGrip;
    ActivateRelease := tmpActivateRelease;
END_IF;

END_FUNCTION_BLOCK

(* ---- public-hard-05.raw_candidate_03.st ---- *)
(* ENGINEERING_CONTRACT
Manual: moving/grip/release outputs are combinational from corresponding button AND NOT corresponding limit switch; releasing the button clears the output. PUB001, PUB005.
SingleStep: rising Start advances only when idle or current step limit reached; each step holds its output until its limit, then waits for next Start. After step 8, next Start goes to step 1. PUB002.
SingleCycle: rising Start starts step 1; each step auto-advances on its completion limit, then stops at step 0 after step 8. PUB003.
Continuous: rising Start starts step 1; auto-advances and loops 8->1. PUB004.
EmergencyStop=FALSE forces all outputs FALSE and freezes automatic state changes. No reset is inferred. PUB005.
Completion feedback uses DownLimitSwitch, UpLimitSwitch, LeftLimitSwitch, RightLimitSwitch, GripLimitSwitch, ReleaseLimitSwitch. Unspecified mode-change behavior preserves the automatic step state.
*)
(* CONTRACT_RULES [] *)
FUNCTION_BLOCK FB_MechanicalArmControl
VAR CONSTANT
    cStepDown1 : INT := 1;
    cStepGrip : INT := 2;
    cStepUp1 : INT := 3;
    cStepRight : INT := 4;
    cStepDown2 : INT := 5;
    cStepRelease : INT := 6;
    cStepUp2 : INT := 7;
    cStepLeft : INT := 8;
END_VAR
VAR_INPUT
    ManualMode : BOOL;
    SingleStepMode : BOOL;
    SingleCycleMode : BOOL;
    ContinuousMode : BOOL;
    EmergencyStop : BOOL;
    Start : BOOL;
    DownButton : BOOL;
    UpButton : BOOL;
    LeftButton : BOOL;
    RightButton : BOOL;
    GripButton : BOOL;
    ReleaseButton : BOOL;
    DownLimitSwitch : BOOL;
    UpLimitSwitch : BOOL;
    LeftLimitSwitch : BOOL;
    RightLimitSwitch : BOOL;
    GripLimitSwitch : BOOL;
    ReleaseLimitSwitch : BOOL;
END_VAR
VAR_OUTPUT
    MoveDown : BOOL;
    MoveUp : BOOL;
    MoveLeft : BOOL;
    MoveRight : BOOL;
    ActivateGrip : BOOL;
    ActivateRelease : BOOL;
END_VAR
VAR
    startTrig : R_TRIG;
    sdStep : INT := 0;
    autoStep : INT := 0;
    sdDone : BOOL;
    autoDone : BOOL;
    tmpMoveDown : BOOL;
    tmpMoveUp : BOOL;
    tmpMoveLeft : BOOL;
    tmpMoveRight : BOOL;
    tmpActivateGrip : BOOL;
    tmpActivateRelease : BOOL;
END_VAR

startTrig(CLK := Start);

tmpMoveDown := FALSE;
tmpMoveUp := FALSE;
tmpMoveLeft := FALSE;
tmpMoveRight := FALSE;
tmpActivateGrip := FALSE;
tmpActivateRelease := FALSE;

IF ManualMode THEN
    tmpMoveDown := DownButton AND NOT DownLimitSwitch;
    tmpMoveUp := UpButton AND NOT UpLimitSwitch;
    tmpMoveLeft := LeftButton AND NOT LeftLimitSwitch;
    tmpMoveRight := RightButton AND NOT RightLimitSwitch;
    tmpActivateGrip := GripButton AND NOT GripLimitSwitch;
    tmpActivateRelease := ReleaseButton AND NOT ReleaseLimitSwitch;

ELSIF SingleStepMode THEN
    CASE sdStep OF
        cStepDown1: sdDone := DownLimitSwitch;
        cStepGrip: sdDone := GripLimitSwitch;
        cStepUp1: sdDone := UpLimitSwitch;
        cStepRight: sdDone := RightLimitSwitch;
        cStepDown2: sdDone := DownLimitSwitch;
        cStepRelease: sdDone := ReleaseLimitSwitch;
        cStepUp2: sdDone := UpLimitSwitch;
        cStepLeft: sdDone := LeftLimitSwitch;
    ELSE
        sdDone := TRUE;
    END_CASE;

    IF EmergencyStop AND startTrig.Q AND sdDone THEN
        IF sdStep >= cStepLeft THEN
            sdStep := cStepDown1;
        ELSE
            sdStep := sdStep + 1;
        END_IF;
    END_IF;

    CASE sdStep OF
        cStepDown1: tmpMoveDown := NOT DownLimitSwitch;
        cStepGrip: tmpActivateGrip := NOT GripLimitSwitch;
        cStepUp1: tmpMoveUp := NOT UpLimitSwitch;
        cStepRight: tmpMoveRight := NOT RightLimitSwitch;
        cStepDown2: tmpMoveDown := NOT DownLimitSwitch;
        cStepRelease: tmpActivateRelease := NOT ReleaseLimitSwitch;
        cStepUp2: tmpMoveUp := NOT UpLimitSwitch;
        cStepLeft: tmpMoveLeft := NOT LeftLimitSwitch;
    ELSE
        (* no automatic output *)
    END_CASE;

ELSIF SingleCycleMode OR ContinuousMode THEN
    IF EmergencyStop AND startTrig.Q AND (autoStep = 0) THEN
        autoStep := cStepDown1;
    END_IF;

    CASE autoStep OF
        cStepDown1: autoDone := DownLimitSwitch;
        cStepGrip: autoDone := GripLimitSwitch;
        cStepUp1: autoDone := UpLimitSwitch;
        cStepRight: autoDone := RightLimitSwitch;
        cStepDown2: autoDone := DownLimitSwitch;
        cStepRelease: autoDone := ReleaseLimitSwitch;
        cStepUp2: autoDone := UpLimitSwitch;
        cStepLeft: autoDone := LeftLimitSwitch;
    ELSE
        autoDone := TRUE;
    END_CASE;

    IF EmergencyStop AND (autoStep <> 0) AND autoDone THEN
        IF SingleCycleMode THEN
            IF autoStep < cStepLeft THEN
                autoStep := autoStep + 1;
            ELSE
                autoStep := 0;
            END_IF;
        ELSIF ContinuousMode THEN
            IF autoStep < cStepLeft THEN
                autoStep := autoStep + 1;
            ELSE
                autoStep := cStepDown1;
            END_IF;
        END_IF;
    END_IF;

    CASE autoStep OF
        cStepDown1: tmpMoveDown := NOT DownLimitSwitch;
        cStepGrip: tmpActivateGrip := NOT GripLimitSwitch;
        cStepUp1: tmpMoveUp := NOT UpLimitSwitch;
        cStepRight: tmpMoveRight := NOT RightLimitSwitch;
        cStepDown2: tmpMoveDown := NOT DownLimitSwitch;
        cStepRelease: tmpActivateRelease := NOT ReleaseLimitSwitch;
        cStepUp2: tmpMoveUp := NOT UpLimitSwitch;
        cStepLeft: tmpMoveLeft := NOT LeftLimitSwitch;
    ELSE
        (* idle/no output *)
    END_CASE;

END_IF;

IF NOT EmergencyStop THEN
    MoveDown := FALSE;
    MoveUp := FALSE;
    MoveLeft := FALSE;
    MoveRight := FALSE;
    ActivateGrip := FALSE;
    ActivateRelease := FALSE;
ELSE
    MoveDown := tmpMoveDown;
    MoveUp := tmpMoveUp;
    MoveLeft := tmpMoveLeft;
    MoveRight := tmpMoveRight;
    ActivateGrip := tmpActivateGrip;
    ActivateRelease := tmpActivateRelease;
END_IF;

END_FUNCTION_BLOCK

(* ---- public-hard-05.raw_candidate_04.st ---- *)
(* ENGINEERING_CONTRACT
Manual: moving/grip/release outputs are combinational from corresponding button AND NOT corresponding limit switch; releasing the button clears the output. PUB001, PUB005.
SingleStep: rising Start advances only when idle or current step limit reached; each step holds its output until its limit, then waits for next Start. After step 8, next Start goes to step 1. PUB002.
SingleCycle: rising Start starts step 1; each step auto-advances on its completion limit, then stops at step 0 after step 8. PUB003.
Continuous: rising Start starts step 1; auto-advances and loops 8->1. PUB004.
EmergencyStop=FALSE forces all outputs FALSE and freezes automatic state changes. No reset is inferred. PUB005.
Completion feedback uses DownLimitSwitch, UpLimitSwitch, LeftLimitSwitch, RightLimitSwitch, GripLimitSwitch, ReleaseLimitSwitch. Unspecified mode-change behavior preserves the automatic step state.
*)
(* CONTRACT_RULES [] *)
FUNCTION_BLOCK FB_MechanicalArmControl
VAR_INPUT
    ManualMode : BOOL;
    SingleStepMode : BOOL;
    SingleCycleMode : BOOL;
    ContinuousMode : BOOL;
    EmergencyStop : BOOL;
    Start : BOOL;
    DownButton : BOOL;
    UpButton : BOOL;
    LeftButton : BOOL;
    RightButton : BOOL;
    GripButton : BOOL;
    ReleaseButton : BOOL;
    DownLimitSwitch : BOOL;
    UpLimitSwitch : BOOL;
    LeftLimitSwitch : BOOL;
    RightLimitSwitch : BOOL;
    GripLimitSwitch : BOOL;
    ReleaseLimitSwitch : BOOL;
END_VAR
VAR_OUTPUT
    MoveDown : BOOL;
    MoveUp : BOOL;
    MoveLeft : BOOL;
    MoveRight : BOOL;
    ActivateGrip : BOOL;
    ActivateRelease : BOOL;
END_VAR
VAR
    startTrig : R_TRIG;
    sdStep : INT := 0;
    autoStep : INT := 0;
    sdDone : BOOL;
    autoDone : BOOL;
    tmpMoveDown : BOOL;
    tmpMoveUp : BOOL;
    tmpMoveLeft : BOOL;
    tmpMoveRight : BOOL;
    tmpActivateGrip : BOOL;
    tmpActivateRelease : BOOL;
END_VAR

startTrig(CLK := Start);

tmpMoveDown := FALSE;
tmpMoveUp := FALSE;
tmpMoveLeft := FALSE;
tmpMoveRight := FALSE;
tmpActivateGrip := FALSE;
tmpActivateRelease := FALSE;

IF ManualMode THEN
    tmpMoveDown := DownButton AND NOT DownLimitSwitch;
    tmpMoveUp := UpButton AND NOT UpLimitSwitch;
    tmpMoveLeft := LeftButton AND NOT LeftLimitSwitch;
    tmpMoveRight := RightButton AND NOT RightLimitSwitch;
    tmpActivateGrip := GripButton AND NOT GripLimitSwitch;
    tmpActivateRelease := ReleaseButton AND NOT ReleaseLimitSwitch;

ELSIF SingleStepMode THEN
    CASE sdStep OF
        1: sdDone := DownLimitSwitch;
        2: sdDone := GripLimitSwitch;
        3: sdDone := UpLimitSwitch;
        4: sdDone := RightLimitSwitch;
        5: sdDone := DownLimitSwitch;
        6: sdDone := ReleaseLimitSwitch;
        7: sdDone := UpLimitSwitch;
        8: sdDone := LeftLimitSwitch;
    ELSE
        sdDone := TRUE;
    END_CASE;

    IF EmergencyStop AND startTrig.Q AND sdDone THEN
        IF sdStep >= 8 THEN
            sdStep := 1;
        ELSE
            sdStep := sdStep + 1;
        END_IF;
    END_IF;

    CASE sdStep OF
        1: tmpMoveDown := NOT DownLimitSwitch;
        2: tmpActivateGrip := NOT GripLimitSwitch;
        3: tmpMoveUp := NOT UpLimitSwitch;
        4: tmpMoveRight := NOT RightLimitSwitch;
        5: tmpMoveDown := NOT DownLimitSwitch;
        6: tmpActivateRelease := NOT ReleaseLimitSwitch;
        7: tmpMoveUp := NOT UpLimitSwitch;
        8: tmpMoveLeft := NOT LeftLimitSwitch;
    END_CASE;

ELSIF (SingleCycleMode OR ContinuousMode) THEN
    IF EmergencyStop AND startTrig.Q AND (autoStep = 0) THEN
        autoStep := 1;
    END_IF;

    CASE autoStep OF
        1: autoDone := DownLimitSwitch;
        2: autoDone := GripLimitSwitch;
        3: autoDone := UpLimitSwitch;
        4: autoDone := RightLimitSwitch;
        5: autoDone := DownLimitSwitch;
        6: autoDone := ReleaseLimitSwitch;
        7: autoDone := UpLimitSwitch;
        8: autoDone := LeftLimitSwitch;
    ELSE
        autoDone := TRUE;
    END_CASE;

    IF EmergencyStop AND (autoStep <> 0) AND autoDone THEN
        IF SingleCycleMode THEN
            IF autoStep < 8 THEN
                autoStep := autoStep + 1;
            ELSE
                autoStep := 0;
            END_IF;
        ELSIF ContinuousMode THEN
            IF autoStep < 8 THEN
                autoStep := autoStep + 1;
            ELSE
                autoStep := 1;
            END_IF;
        END_IF;
    END_IF;

    CASE autoStep OF
        1: tmpMoveDown := NOT DownLimitSwitch;
        2: tmpActivateGrip := NOT GripLimitSwitch;
        3: tmpMoveUp := NOT UpLimitSwitch;
        4: tmpMoveRight := NOT RightLimitSwitch;
        5: tmpMoveDown := NOT DownLimitSwitch;
        6: tmpActivateRelease := NOT ReleaseLimitSwitch;
        7: tmpMoveUp := NOT UpLimitSwitch;
        8: tmpMoveLeft := NOT LeftLimitSwitch;
    END_CASE;

END_IF;

IF NOT EmergencyStop THEN
    MoveDown := FALSE;
    MoveUp := FALSE;
    MoveLeft := FALSE;
    MoveRight := FALSE;
    ActivateGrip := FALSE;
    ActivateRelease := FALSE;
ELSE
    MoveDown := tmpMoveDown;
    MoveUp := tmpMoveUp;
    MoveLeft := tmpMoveLeft;
    MoveRight := tmpMoveRight;
    ActivateGrip := tmpActivateGrip;
    ActivateRelease := tmpActivateRelease;
END_IF;

END_FUNCTION_BLOCK

(* ---- public-hard-06.candidate_01.st ---- *)
(* ENGINEERING_CONTRACT
MotorForward (auto): activated by state machine transfer legs PUB003/PUB004; held while state; off at target sensor or manual PUB002.
MotorForward (manual): ForwardButton level, interlocked; PUB002.
MotorReverse (manual): ReverseButton level, interlocked; both buttons -> both off.
kick: unqualified after weightComplete at weighing; latched until SensorWeight false (unspecified removal); PUB004.
CompletionLight: on at SensorOutput arrival after firing, held until SensorOutput false; PUB004.
firingTemp: linear 100->500, 200->550 inclusive; set on qualified weighing; retained otherwise; PUB004.
State localState: retained across scans; mode switch does not reset; unspecified reset on mode change.
*)
(* CONTRACT_RULES [] *)
TYPE ProductionLineState :
(
    STATE_IDLE,
    STATE_MOVING_TO_WASH,
    STATE_AT_WASH,
    STATE_MOVING_TO_WEIGH,
    STATE_AT_WEIGH,
    STATE_MOVING_TO_FIRING,
    STATE_AT_FIRING,
    STATE_MOVING_TO_OUTPUT,
    STATE_AT_OUTPUT
);
END_TYPE;

FUNCTION_BLOCK ProductionControl
VAR_INPUT
    Mode : BOOL;
    ForwardButton : BOOL;
    ReverseButton : BOOL;
    SensorFeed : BOOL;
    SensorWash : BOOL;
    SensorWeight : BOOL;
    SensorFiring : BOOL;
    SensorOutput : BOOL;
    washComplete : BOOL;
    weightComplete : BOOL;
    weight : REAL;
    firingComplete : BOOL;
END_VAR
VAR_OUTPUT
    MotorForward : BOOL;
    MotorReverse : BOOL;
    kick : BOOL;
    CompletionLight : BOOL;
    firingTemp : REAL;
END_VAR
VAR
    localState : ProductionLineState := STATE_IDLE;
    localKickActive : BOOL := FALSE;
END_VAR

IF Mode THEN
    MotorReverse := FALSE;

    CASE localState OF
        STATE_IDLE:
            MotorForward := FALSE;
            CompletionLight := FALSE;
            kick := FALSE;
            localKickActive := FALSE;
            IF SensorFeed THEN
                MotorForward := TRUE;
                localState := STATE_MOVING_TO_WASH;
            END_IF;

        STATE_MOVING_TO_WASH:
            MotorForward := TRUE;
            IF SensorWash THEN
                MotorForward := FALSE;
                localState := STATE_AT_WASH;
            END_IF;

        STATE_AT_WASH:
            MotorForward := FALSE;
            IF washComplete THEN
                MotorForward := TRUE;
                localState := STATE_MOVING_TO_WEIGH;
            END_IF;

        STATE_MOVING_TO_WEIGH:
            MotorForward := TRUE;
            IF SensorWeight THEN
                MotorForward := FALSE;
                localState := STATE_AT_WEIGH;
            END_IF;

        STATE_AT_WEIGH:
            MotorForward := FALSE;
            IF localKickActive THEN
                IF NOT SensorWeight THEN
                    kick := FALSE;
                    localKickActive := FALSE;
                    localState := STATE_IDLE;
                END_IF;
            ELSIF weightComplete THEN
                IF (weight >= 100.0) AND (weight <= 200.0) THEN
                    firingTemp := 500.0 + (weight - 100.0) * 0.5;
                    kick := FALSE;
                    localKickActive := FALSE;
                    MotorForward := TRUE;
                    localState := STATE_MOVING_TO_FIRING;
                ELSE
                    kick := TRUE;
                    localKickActive := TRUE;
                    MotorForward := FALSE;
                END_IF;
            END_IF;

        STATE_MOVING_TO_FIRING:
            MotorForward := TRUE;
            IF SensorFiring THEN
                MotorForward := FALSE;
                localState := STATE_AT_FIRING;
            END_IF;

        STATE_AT_FIRING:
            MotorForward := FALSE;
            IF firingComplete THEN
                MotorForward := TRUE;
                localState := STATE_MOVING_TO_OUTPUT;
            END_IF;

        STATE_MOVING_TO_OUTPUT:
            MotorForward := TRUE;
            CompletionLight := FALSE;
            IF SensorOutput THEN
                MotorForward := FALSE;
                CompletionLight := TRUE;
                localState := STATE_AT_OUTPUT;
            END_IF;

        STATE_AT_OUTPUT:
            MotorForward := FALSE;
            CompletionLight := TRUE;
            IF NOT SensorOutput THEN
                CompletionLight := FALSE;
                localState := STATE_IDLE;
            END_IF;
    END_CASE;

ELSE
    MotorForward := ForwardButton AND (NOT ReverseButton);
    MotorReverse := ReverseButton AND (NOT ForwardButton);
    (* kick, CompletionLight, firingTemp retain their last automatic values *)
END_IF;

END_FUNCTION_BLOCK

(* ---- public-hard-06.candidate_02.st ---- *)
(* ENGINEERING_CONTRACT
MotorForward (auto): activated by state machine transfer legs PUB003/PUB004; held while state; off at target sensor or manual PUB002.
MotorForward (manual): ForwardButton level, interlocked; PUB002.
MotorReverse (manual): ReverseButton level, interlocked; both buttons -> both off.
kick: unqualified after weightComplete at weighing; latched until SensorWeight false (unspecified removal); PUB004.
CompletionLight: on at SensorOutput arrival after firing, held until SensorOutput false; PUB004.
firingTemp: linear 100->500, 200->550 inclusive; set on qualified weighing; retained otherwise; PUB004.
State localState: retained across scans; manual mode resets automatic sequence to IDLE; unspecified otherwise.
*)
(* CONTRACT_RULES [] *)
TYPE ProductionLineState :
(
    STATE_IDLE,
    STATE_MOVING_TO_WASH,
    STATE_AT_WASH,
    STATE_MOVING_TO_WEIGH,
    STATE_AT_WEIGH,
    STATE_MOVING_TO_FIRING,
    STATE_AT_FIRING,
    STATE_MOVING_TO_OUTPUT,
    STATE_AT_OUTPUT
);
END_TYPE;

FUNCTION_BLOCK ProductionControl
VAR_INPUT
    Mode : BOOL;
    ForwardButton : BOOL;
    ReverseButton : BOOL;
    SensorFeed : BOOL;
    SensorWash : BOOL;
    SensorWeight : BOOL;
    SensorFiring : BOOL;
    SensorOutput : BOOL;
    washComplete : BOOL;
    weightComplete : BOOL;
    weight : REAL;
    firingComplete : BOOL;
END_VAR
VAR_OUTPUT
    MotorForward : BOOL;
    MotorReverse : BOOL;
    kick : BOOL;
    CompletionLight : BOOL;
    firingTemp : REAL;
END_VAR
VAR
    localState : ProductionLineState := STATE_IDLE;
    localKickActive : BOOL := FALSE;
END_VAR

IF Mode THEN
    MotorReverse := FALSE;

    CASE localState OF
        STATE_IDLE:
            MotorForward := FALSE;
            CompletionLight := FALSE;
            kick := FALSE;
            localKickActive := FALSE;
            IF SensorFeed THEN
                MotorForward := TRUE;
                localState := STATE_MOVING_TO_WASH;
            END_IF;

        STATE_MOVING_TO_WASH:
            MotorForward := TRUE;
            IF SensorWash THEN
                MotorForward := FALSE;
                localState := STATE_AT_WASH;
            END_IF;

        STATE_AT_WASH:
            MotorForward := FALSE;
            IF washComplete THEN
                MotorForward := TRUE;
                localState := STATE_MOVING_TO_WEIGH;
            END_IF;

        STATE_MOVING_TO_WEIGH:
            MotorForward := TRUE;
            IF SensorWeight THEN
                MotorForward := FALSE;
                localState := STATE_AT_WEIGH;
            END_IF;

        STATE_AT_WEIGH:
            MotorForward := FALSE;
            IF localKickActive THEN
                IF NOT SensorWeight THEN
                    kick := FALSE;
                    localKickActive := FALSE;
                    localState := STATE_IDLE;
                END_IF;
            ELSIF weightComplete THEN
                IF (weight >= 100.0) AND (weight <= 200.0) THEN
                    firingTemp := 500.0 + (weight - 100.0) * 0.5;
                    kick := FALSE;
                    localKickActive := FALSE;
                    MotorForward := TRUE;
                    localState := STATE_MOVING_TO_FIRING;
                ELSE
                    kick := TRUE;
                    localKickActive := TRUE;
                    MotorForward := FALSE;
                END_IF;
            END_IF;

        STATE_MOVING_TO_FIRING:
            MotorForward := TRUE;
            IF SensorFiring THEN
                MotorForward := FALSE;
                localState := STATE_AT_FIRING;
            END_IF;

        STATE_AT_FIRING:
            MotorForward := FALSE;
            IF firingComplete THEN
                MotorForward := TRUE;
                localState := STATE_MOVING_TO_OUTPUT;
            END_IF;

        STATE_MOVING_TO_OUTPUT:
            MotorForward := TRUE;
            CompletionLight := FALSE;
            IF SensorOutput THEN
                MotorForward := FALSE;
                CompletionLight := TRUE;
                localState := STATE_AT_OUTPUT;
            END_IF;

        STATE_AT_OUTPUT:
            MotorForward := FALSE;
            CompletionLight := TRUE;
            IF NOT SensorOutput THEN
                CompletionLight := FALSE;
                localState := STATE_IDLE;
            END_IF;
    END_CASE;

ELSE
    MotorForward := ForwardButton AND (NOT ReverseButton);
    MotorReverse := ReverseButton AND (NOT ForwardButton);
    localState := STATE_IDLE;
    localKickActive := FALSE;
    (* kick, CompletionLight, firingTemp retain their last automatic values *)
END_IF;

END_FUNCTION_BLOCK

(* ---- public-hard-06.raw_candidate_01.st ---- *)
(* ENGINEERING_CONTRACT
MotorForward (auto): activated by state machine transfer legs PUB003/PUB004; held while state; off at target sensor or manual PUB002.
MotorForward (manual): ForwardButton level, interlocked; PUB002.
MotorReverse (manual): ReverseButton level, interlocked; both buttons -> both off.
kick: unqualified after weightComplete at weighing; latched until SensorWeight false (unspecified removal); PUB004.
CompletionLight: on at SensorOutput arrival after firing, held until SensorOutput false; PUB004.
firingTemp: linear 100->500, 200->550 inclusive; set on qualified weighing; retained otherwise; PUB004.
State localState: retained across scans; mode switch does not reset; unspecified reset on mode change.
*)
(* CONTRACT_RULES [] *)
TYPE ProductionLineState :
(
    STATE_IDLE,
    STATE_MOVING_TO_WASH,
    STATE_AT_WASH,
    STATE_MOVING_TO_WEIGH,
    STATE_AT_WEIGH,
    STATE_MOVING_TO_FIRING,
    STATE_AT_FIRING,
    STATE_MOVING_TO_OUTPUT,
    STATE_AT_OUTPUT
);
END_TYPE

FUNCTION_BLOCK ProductionControl
VAR_INPUT
    Mode : BOOL;
    ForwardButton : BOOL;
    ReverseButton : BOOL;
    SensorFeed : BOOL;
    SensorWash : BOOL;
    SensorWeight : BOOL;
    SensorFiring : BOOL;
    SensorOutput : BOOL;
    washComplete : BOOL;
    weightComplete : BOOL;
    weight : REAL;
    firingComplete : BOOL;
END_VAR
VAR_OUTPUT
    MotorForward : BOOL;
    MotorReverse : BOOL;
    kick : BOOL;
    CompletionLight : BOOL;
    firingTemp : REAL;
END_VAR
VAR
    localState : ProductionLineState := STATE_IDLE;
    localKickActive : BOOL := FALSE;
END_VAR

IF Mode THEN
    MotorReverse := FALSE;

    CASE localState OF
        STATE_IDLE:
            MotorForward := FALSE;
            CompletionLight := FALSE;
            kick := FALSE;
            localKickActive := FALSE;
            IF SensorFeed THEN
                MotorForward := TRUE;
                localState := STATE_MOVING_TO_WASH;
            END_IF;

        STATE_MOVING_TO_WASH:
            MotorForward := TRUE;
            IF SensorWash THEN
                MotorForward := FALSE;
                localState := STATE_AT_WASH;
            END_IF;

        STATE_AT_WASH:
            MotorForward := FALSE;
            IF washComplete THEN
                MotorForward := TRUE;
                localState := STATE_MOVING_TO_WEIGH;
            END_IF;

        STATE_MOVING_TO_WEIGH:
            MotorForward := TRUE;
            IF SensorWeight THEN
                MotorForward := FALSE;
                localState := STATE_AT_WEIGH;
            END_IF;

        STATE_AT_WEIGH:
            MotorForward := FALSE;
            IF localKickActive THEN
                IF NOT SensorWeight THEN
                    kick := FALSE;
                    localKickActive := FALSE;
                    localState := STATE_IDLE;
                END_IF;
            ELSIF weightComplete THEN
                IF (weight >= 100.0) AND (weight <= 200.0) THEN
                    firingTemp := 500.0 + (weight - 100.0) * 0.5;
                    kick := FALSE;
                    localKickActive := FALSE;
                    MotorForward := TRUE;
                    localState := STATE_MOVING_TO_FIRING;
                ELSE
                    kick := TRUE;
                    localKickActive := TRUE;
                    MotorForward := FALSE;
                END_IF;
            END_IF;

        STATE_MOVING_TO_FIRING:
            MotorForward := TRUE;
            IF SensorFiring THEN
                MotorForward := FALSE;
                localState := STATE_AT_FIRING;
            END_IF;

        STATE_AT_FIRING:
            MotorForward := FALSE;
            IF firingComplete THEN
                MotorForward := TRUE;
                localState := STATE_MOVING_TO_OUTPUT;
            END_IF;

        STATE_MOVING_TO_OUTPUT:
            MotorForward := TRUE;
            CompletionLight := FALSE;
            IF SensorOutput THEN
                MotorForward := FALSE;
                CompletionLight := TRUE;
                localState := STATE_AT_OUTPUT;
            END_IF;

        STATE_AT_OUTPUT:
            MotorForward := FALSE;
            CompletionLight := TRUE;
            IF NOT SensorOutput THEN
                CompletionLight := FALSE;
                localState := STATE_IDLE;
            END_IF;
    END_CASE;

ELSE
    MotorForward := ForwardButton AND (NOT ReverseButton);
    MotorReverse := ReverseButton AND (NOT ForwardButton);
    (* kick, CompletionLight, firingTemp retain their last automatic values *)
END_IF;

END_FUNCTION_BLOCK

(* ---- public-hard-06.raw_candidate_02.st ---- *)
(* ENGINEERING_CONTRACT
MotorForward (auto): activated by state machine transfer legs PUB003/PUB004; held while state; off at target sensor or manual PUB002.
MotorForward (manual): ForwardButton level, interlocked; PUB002.
MotorReverse (manual): ReverseButton level, interlocked; both buttons -> both off.
kick: unqualified after weightComplete at weighing; latched until SensorWeight false (unspecified removal); PUB004.
CompletionLight: on at SensorOutput arrival after firing, held until SensorOutput false; PUB004.
firingTemp: linear 100->500, 200->550 inclusive; set on qualified weighing; retained otherwise; PUB004.
State localState: retained across scans; manual mode resets automatic sequence to IDLE; unspecified otherwise.
*)
(* CONTRACT_RULES [] *)
TYPE ProductionLineState :
(
    STATE_IDLE,
    STATE_MOVING_TO_WASH,
    STATE_AT_WASH,
    STATE_MOVING_TO_WEIGH,
    STATE_AT_WEIGH,
    STATE_MOVING_TO_FIRING,
    STATE_AT_FIRING,
    STATE_MOVING_TO_OUTPUT,
    STATE_AT_OUTPUT
);
END_TYPE;

FUNCTION_BLOCK ProductionControl
VAR_INPUT
    Mode : BOOL;
    ForwardButton : BOOL;
    ReverseButton : BOOL;
    SensorFeed : BOOL;
    SensorWash : BOOL;
    SensorWeight : BOOL;
    SensorFiring : BOOL;
    SensorOutput : BOOL;
    washComplete : BOOL;
    weightComplete : BOOL;
    weight : REAL;
    firingComplete : BOOL;
END_VAR
VAR_OUTPUT
    MotorForward : BOOL;
    MotorReverse : BOOL;
    kick : BOOL;
    CompletionLight : BOOL;
    firingTemp : REAL;
END_VAR
VAR
    localState : ProductionLineState := STATE_IDLE;
    localKickActive : BOOL := FALSE;
END_VAR

IF Mode THEN
    MotorReverse := FALSE;

    CASE localState OF
        STATE_IDLE:
            MotorForward := FALSE;
            CompletionLight := FALSE;
            kick := FALSE;
            localKickActive := FALSE;
            IF SensorFeed THEN
                MotorForward := TRUE;
                localState := STATE_MOVING_TO_WASH;
            END_IF;

        STATE_MOVING_TO_WASH:
            MotorForward := TRUE;
            IF SensorWash THEN
                MotorForward := FALSE;
                localState := STATE_AT_WASH;
            END_IF;

        STATE_AT_WASH:
            MotorForward := FALSE;
            IF washComplete THEN
                MotorForward := TRUE;
                localState := STATE_MOVING_TO_WEIGH;
            END_IF;

        STATE_MOVING_TO_WEIGH:
            MotorForward := TRUE;
            IF SensorWeight THEN
                MotorForward := FALSE;
                localState := STATE_AT_WEIGH;
            END_IF;

        STATE_AT_WEIGH:
            MotorForward := FALSE;
            IF localKickActive THEN
                IF NOT SensorWeight THEN
                    kick := FALSE;
                    localKickActive := FALSE;
                    localState := STATE_IDLE;
                END_IF;
            ELSIF weightComplete THEN
                IF (weight >= 100.0) AND (weight <= 200.0) THEN
                    firingTemp := 500.0 + (weight - 100.0) * 0.5;
                    kick := FALSE;
                    localKickActive := FALSE;
                    MotorForward := TRUE;
                    localState := STATE_MOVING_TO_FIRING;
                ELSE
                    kick := TRUE;
                    localKickActive := TRUE;
                    MotorForward := FALSE;
                END_IF;
            END_IF;

        STATE_MOVING_TO_FIRING:
            MotorForward := TRUE;
            IF SensorFiring THEN
                MotorForward := FALSE;
                localState := STATE_AT_FIRING;
            END_IF;

        STATE_AT_FIRING:
            MotorForward := FALSE;
            IF firingComplete THEN
                MotorForward := TRUE;
                localState := STATE_MOVING_TO_OUTPUT;
            END_IF;

        STATE_MOVING_TO_OUTPUT:
            MotorForward := TRUE;
            CompletionLight := FALSE;
            IF SensorOutput THEN
                MotorForward := FALSE;
                CompletionLight := TRUE;
                localState := STATE_AT_OUTPUT;
            END_IF;

        STATE_AT_OUTPUT:
            MotorForward := FALSE;
            CompletionLight := TRUE;
            IF NOT SensorOutput THEN
                CompletionLight := FALSE;
                localState := STATE_IDLE;
            END_IF;
    END_CASE;

ELSE
    MotorForward := ForwardButton AND (NOT ReverseButton);
    MotorReverse := ReverseButton AND (NOT ForwardButton);
    localState := STATE_IDLE;
    localKickActive := FALSE;
    (* kick, CompletionLight, firingTemp retain their last automatic values *)
END_IF;

END_FUNCTION_BLOCK

(* ---- public-medium-01.candidate_01.st ---- *)
(* ENGINEERING_CONTRACT
   - Mode FALSE=manual, TRUE=automatic (PUB001).
   - Latched local_Running: start sets TRUE, stop clears; same-scan stop wins (PUB002).
   - When local_Running=FALSE, all RunComd are FALSE (PUB002).
   - Manual and running: each RunComd follows its current selection each scan (PUB001).
   - Automatic and running: select 3 highest priority pumps, larger priority wins;
     ties are resolved to the lowest array index; remaining two are stopped (PUB003).
   - priority and selection are read-only; only RunComd is written (PUB004).
   - Unspecified: initial state is stopped; priority/selection changes take effect while Running.
*)
(* CONTRACT_RULES [] *)
TYPE ST_Pump :
STRUCT
    priority : INT;
    selection : BOOL;
    RunComd : BOOL;
END_STRUCT
END_TYPE;

FUNCTION_BLOCK FB_MultiPumpControl
VAR_INPUT
    mode : BOOL;
    start : BOOL;
    stop : BOOL;
END_VAR
VAR_IN_OUT
    pumpGroup : ARRAY[1..5] OF ST_Pump;
END_VAR
VAR
    local_Running : BOOL;
    local_selected : ARRAY[1..5] OF BOOL;
    local_bestIdx : INT;
    local_bestPrio : INT;
    local_i : INT;
    local_j : INT;
END_VAR

IF stop THEN
    local_Running := FALSE;
ELSIF start THEN
    local_Running := TRUE;
END_IF;

IF NOT local_Running THEN
    FOR local_i := 1 TO 5 DO
        pumpGroup[local_i].RunComd := FALSE;
    END_FOR;
ELSE
    IF NOT mode THEN
        FOR local_i := 1 TO 5 DO
            pumpGroup[local_i].RunComd := pumpGroup[local_i].selection;
        END_FOR;
    ELSE
        FOR local_i := 1 TO 5 DO
            local_selected[local_i] := FALSE;
        END_FOR;

        FOR local_j := 1 TO 3 DO
            local_bestIdx := 0;
            local_bestPrio := -32768;

            FOR local_i := 1 TO 5 DO
                IF NOT local_selected[local_i] THEN
                    IF (local_bestIdx = 0) OR (pumpGroup[local_i].priority > local_bestPrio) THEN
                        local_bestIdx := local_i;
                        local_bestPrio := pumpGroup[local_i].priority;
                    END_IF;
                END_IF;
            END_FOR;

            IF local_bestIdx <> 0 THEN
                local_selected[local_bestIdx] := TRUE;
            END_IF;
        END_FOR;

        FOR local_i := 1 TO 5 DO
            pumpGroup[local_i].RunComd := local_selected[local_i];
        END_FOR;
    END_IF;
END_IF;

END_FUNCTION_BLOCK

(* ---- public-medium-01.candidate_02.st ---- *)
(* ENGINEERING_CONTRACT
   - Mode FALSE=manual, TRUE=automatic (PUB001).
   - start is rising-edge triggered; stop is level-sensitive with priority (PUB002).
   - Latched local_Running: start edge sets TRUE; stop clears; stop wins (PUB002).
   - When local_Running=FALSE, all RunComd are FALSE (PUB002).
   - Manual and running: each RunComd follows its current selection each scan (PUB001).
   - Automatic and running: select 3 highest priority pumps, larger priority wins;
     ties resolved to lowest array index; remaining two stopped (PUB003).
   - priority and selection are read-only; only RunComd written (PUB004).
   - Unspecified: initial state stopped; priority/selection changes take effect while Running.
*)
(* CONTRACT_RULES [] *)
TYPE ST_Pump :
STRUCT
    priority : INT;
    selection : BOOL;
    RunComd : BOOL;
END_STRUCT
END_TYPE;

FUNCTION_BLOCK FB_MultiPumpControl
VAR_INPUT
    mode : BOOL;
    start : BOOL;
    stop : BOOL;
END_VAR
VAR_IN_OUT
    pumpGroup : ARRAY[1..5] OF ST_Pump;
END_VAR
VAR
    local_Running : BOOL;
    local_start_prev : BOOL;
    local_start_rising : BOOL;
    local_selected : ARRAY[1..5] OF BOOL;
    local_bestIdx : INT;
    local_bestPrio : INT;
    local_i : INT;
    local_j : INT;
END_VAR

(* Detect rising edge of start *)
local_start_rising := start AND NOT local_start_prev;

IF stop THEN
    local_Running := FALSE;
ELSIF local_start_rising THEN
    local_Running := TRUE;
END_IF;

(* Update start previous state for next scan *)
local_start_prev := start;

IF NOT local_Running THEN
    FOR local_i := 1 TO 5 DO
        pumpGroup[local_i].RunComd := FALSE;
    END_FOR;
ELSE
    IF NOT mode THEN
        FOR local_i := 1 TO 5 DO
            pumpGroup[local_i].RunComd := pumpGroup[local_i].selection;
        END_FOR;
    ELSE
        FOR local_i := 1 TO 5 DO
            local_selected[local_i] := FALSE;
        END_FOR;

        FOR local_j := 1 TO 3 DO
            local_bestIdx := 0;
            local_bestPrio := -32768;

            FOR local_i := 1 TO 5 DO
                IF NOT local_selected[local_i] THEN
                    IF (local_bestIdx = 0) OR (pumpGroup[local_i].priority > local_bestPrio) THEN
                        local_bestIdx := local_i;
                        local_bestPrio := pumpGroup[local_i].priority;
                    END_IF;
                END_IF;
            END_FOR;

            IF local_bestIdx <> 0 THEN
                local_selected[local_bestIdx] := TRUE;
            END_IF;
        END_FOR;

        FOR local_i := 1 TO 5 DO
            pumpGroup[local_i].RunComd := local_selected[local_i];
        END_FOR;
    END_IF;
END_IF;

END_FUNCTION_BLOCK

(* ---- public-medium-01.candidate_03.st ---- *)
(* ENGINEERING_CONTRACT
   - Mode FALSE=manual, TRUE=automatic (PUB001).
   - local_Running is retained run command: set by start OR previous running, cleared by stop; stop level wins (PUB002).
   - When local_Running=FALSE, all RunComd are FALSE (PUB002).
   - Manual running: each RunComd follows its current selection each scan (PUB001).
   - Automatic running: select 3 highest priority pumps, tie lower index; remaining stopped (PUB003).
   - priority/selection read-only; only RunComd written (PUB004).
*)
(* CONTRACT_RULES [] *)
TYPE ST_Pump :
STRUCT
    priority : INT;
    selection : BOOL;
    RunComd : BOOL;
END_STRUCT
END_TYPE;

FUNCTION_BLOCK FB_MultiPumpControl
VAR_INPUT
    mode : BOOL;
    start : BOOL;
    stop : BOOL;
END_VAR
VAR_IN_OUT
    pumpGroup : ARRAY[1..5] OF ST_Pump;
END_VAR
VAR
    local_Running : BOOL;
    local_selected : ARRAY[1..5] OF BOOL;
    local_bestIdx : INT;
    local_bestPrio : INT;
    local_i : INT;
    local_j : INT;
END_VAR

IF stop THEN
    local_Running := FALSE;
ELSE
    local_Running := local_Running OR start;
END_IF;

IF NOT local_Running THEN
    FOR local_i := 1 TO 5 DO
        pumpGroup[local_i].RunComd := FALSE;
    END_FOR;
ELSE
    IF NOT mode THEN
        FOR local_i := 1 TO 5 DO
            pumpGroup[local_i].RunComd := pumpGroup[local_i].selection;
        END_FOR;
    ELSE
        FOR local_i := 1 TO 5 DO
            local_selected[local_i] := FALSE;
        END_FOR;

        FOR local_j := 1 TO 3 DO
            local_bestIdx := 0;
            local_bestPrio := -32768;

            FOR local_i := 1 TO 5 DO
                IF NOT local_selected[local_i] THEN
                    IF (local_bestIdx = 0) OR (pumpGroup[local_i].priority > local_bestPrio) THEN
                        local_bestIdx := local_i;
                        local_bestPrio := pumpGroup[local_i].priority;
                    END_IF;
                END_IF;
            END_FOR;

            IF local_bestIdx <> 0 THEN
                local_selected[local_bestIdx] := TRUE;
            END_IF;
        END_FOR;

        FOR local_i := 1 TO 5 DO
            pumpGroup[local_i].RunComd := local_selected[local_i];
        END_FOR;
    END_IF;
END_IF;

END_FUNCTION_BLOCK

(* ---- public-medium-01.candidate_04.st ---- *)
(* ENGINEERING_CONTRACT
   - Mode FALSE=manual, TRUE=automatic (PUB001).
   - Start is edge-triggered: a new FALSE->TRUE start pulse is required after stop release
     before pumps may run again; stop has priority over a level-held start (PUB001/PUB002).
   - local_Running is retained run state: set by rising edge of start while stop=FALSE,
     cleared immediately by stop=TRUE (PUB002).
   - When local_Running=FALSE, all RunComd are FALSE (PUB002).
   - Manual running: each RunComd follows its current selection each scan (PUB001).
   - Automatic running: select 3 highest priority pumps, tie lower index; remaining stopped (PUB003).
   - priority/selection read-only; only RunComd written (PUB004).
*)
(* CONTRACT_RULES [] *)
TYPE ST_Pump :
STRUCT
    priority : INT;
    selection : BOOL;
    RunComd : BOOL;
END_STRUCT
END_TYPE;

FUNCTION_BLOCK FB_MultiPumpControl
VAR_INPUT
    mode : BOOL;
    start : BOOL;
    stop : BOOL;
END_VAR
VAR_IN_OUT
    pumpGroup : ARRAY[1..5] OF ST_Pump;
END_VAR
VAR
    local_Running : BOOL;
    local_selected : ARRAY[1..5] OF BOOL;
    local_bestIdx : INT;
    local_bestPrio : INT;
    local_i : INT;
    local_j : INT;
    local_rtStart : R_TRIG;
END_VAR

local_rtStart(CLK := start);

IF stop THEN
    local_Running := FALSE;
ELSE
    local_Running := local_Running OR local_rtStart.Q;
END_IF;

IF NOT local_Running THEN
    FOR local_i := 1 TO 5 DO
        pumpGroup[local_i].RunComd := FALSE;
    END_FOR;
ELSE
    IF NOT mode THEN
        FOR local_i := 1 TO 5 DO
            pumpGroup[local_i].RunComd := pumpGroup[local_i].selection;
        END_FOR;
    ELSE
        FOR local_i := 1 TO 5 DO
            local_selected[local_i] := FALSE;
        END_FOR;

        FOR local_j := 1 TO 3 DO
            local_bestIdx := 0;
            local_bestPrio := -32768;

            FOR local_i := 1 TO 5 DO
                IF NOT local_selected[local_i] THEN
                    IF (local_bestIdx = 0) OR (pumpGroup[local_i].priority > local_bestPrio) THEN
                        local_bestIdx := local_i;
                        local_bestPrio := pumpGroup[local_i].priority;
                    END_IF;
                END_IF;
            END_FOR;

            IF local_bestIdx <> 0 THEN
                local_selected[local_bestIdx] := TRUE;
            END_IF;
        END_FOR;

        FOR local_i := 1 TO 5 DO
            pumpGroup[local_i].RunComd := local_selected[local_i];
        END_FOR;
    END_IF;
END_IF;

END_FUNCTION_BLOCK

(* ---- public-medium-01.raw_candidate_01.st ---- *)
(* ENGINEERING_CONTRACT
   - Mode FALSE=manual, TRUE=automatic (PUB001).
   - Latched local_Running: start sets TRUE, stop clears; same-scan stop wins (PUB002).
   - When local_Running=FALSE, all RunComd are FALSE (PUB002).
   - Manual and running: each RunComd follows its current selection each scan (PUB001).
   - Automatic and running: select 3 highest priority pumps, larger priority wins;
     ties are resolved to the lowest array index; remaining two are stopped (PUB003).
   - priority and selection are read-only; only RunComd is written (PUB004).
   - Unspecified: initial state is stopped; priority/selection changes take effect while Running.
*)
(* CONTRACT_RULES [] *)
TYPE ST_Pump :
STRUCT
    priority : INT;
    selection : BOOL;
    RunComd : BOOL;
END_STRUCT
END_TYPE

FUNCTION_BLOCK FB_MultiPumpControl
VAR_INPUT
    mode : BOOL;
    start : BOOL;
    stop : BOOL;
END_VAR
VAR_IN_OUT
    pumpGroup : ARRAY[1..5] OF ST_Pump;
END_VAR
VAR
    local_Running : BOOL;
    local_selected : ARRAY[1..5] OF BOOL;
    local_bestIdx : INT;
    local_bestPrio : INT;
    local_i : INT;
    local_j : INT;
END_VAR

IF stop THEN
    local_Running := FALSE;
ELSIF start THEN
    local_Running := TRUE;
END_IF;

IF NOT local_Running THEN
    FOR local_i := 1 TO 5 DO
        pumpGroup[local_i].RunComd := FALSE;
    END_FOR;
ELSE
    IF NOT mode THEN
        FOR local_i := 1 TO 5 DO
            pumpGroup[local_i].RunComd := pumpGroup[local_i].selection;
        END_FOR;
    ELSE
        FOR local_i := 1 TO 5 DO
            local_selected[local_i] := FALSE;
        END_FOR;

        FOR local_j := 1 TO 3 DO
            local_bestIdx := 0;
            local_bestPrio := -32768;

            FOR local_i := 1 TO 5 DO
                IF NOT local_selected[local_i] THEN
                    IF (local_bestIdx = 0) OR (pumpGroup[local_i].priority > local_bestPrio) THEN
                        local_bestIdx := local_i;
                        local_bestPrio := pumpGroup[local_i].priority;
                    END_IF;
                END_IF;
            END_FOR;

            IF local_bestIdx <> 0 THEN
                local_selected[local_bestIdx] := TRUE;
            END_IF;
        END_FOR;

        FOR local_i := 1 TO 5 DO
            pumpGroup[local_i].RunComd := local_selected[local_i];
        END_FOR;
    END_IF;
END_IF;

END_FUNCTION_BLOCK

(* ---- public-medium-01.raw_candidate_02.st ---- *)
(* ENGINEERING_CONTRACT
   - Mode FALSE=manual, TRUE=automatic (PUB001).
   - start is rising-edge triggered; stop is level-sensitive with priority (PUB002).
   - Latched local_Running: start edge sets TRUE; stop clears; stop wins (PUB002).
   - When local_Running=FALSE, all RunComd are FALSE (PUB002).
   - Manual and running: each RunComd follows its current selection each scan (PUB001).
   - Automatic and running: select 3 highest priority pumps, larger priority wins;
     ties resolved to lowest array index; remaining two stopped (PUB003).
   - priority and selection are read-only; only RunComd written (PUB004).
   - Unspecified: initial state stopped; priority/selection changes take effect while Running.
*)
(* CONTRACT_RULES [] *)
TYPE ST_Pump :
STRUCT
    priority : INT;
    selection : BOOL;
    RunComd : BOOL;
END_STRUCT
END_TYPE;

FUNCTION_BLOCK FB_MultiPumpControl
VAR_INPUT
    mode : BOOL;
    start : BOOL;
    stop : BOOL;
END_VAR
VAR_IN_OUT
    pumpGroup : ARRAY[1..5] OF ST_Pump;
END_VAR
VAR
    local_Running : BOOL;
    local_start_prev : BOOL;
    local_start_rising : BOOL;
    local_selected : ARRAY[1..5] OF BOOL;
    local_bestIdx : INT;
    local_bestPrio : INT;
    local_i : INT;
    local_j : INT;
END_VAR

(* Detect rising edge of start *)
local_start_rising := start AND NOT local_start_prev;

IF stop THEN
    local_Running := FALSE;
ELSIF local_start_rising THEN
    local_Running := TRUE;
END_IF;

(* Update start previous state for next scan *)
local_start_prev := start;

IF NOT local_Running THEN
    FOR local_i := 1 TO 5 DO
        pumpGroup[local_i].RunComd := FALSE;
    END_FOR;
ELSE
    IF NOT mode THEN
        FOR local_i := 1 TO 5 DO
            pumpGroup[local_i].RunComd := pumpGroup[local_i].selection;
        END_FOR;
    ELSE
        FOR local_i := 1 TO 5 DO
            local_selected[local_i] := FALSE;
        END_FOR;

        FOR local_j := 1 TO 3 DO
            local_bestIdx := 0;
            local_bestPrio := -32768;

            FOR local_i := 1 TO 5 DO
                IF NOT local_selected[local_i] THEN
                    IF (local_bestIdx = 0) OR (pumpGroup[local_i].priority > local_bestPrio) THEN
                        local_bestIdx := local_i;
                        local_bestPrio := pumpGroup[local_i].priority;
                    END_IF;
                END_IF;
            END_FOR;

            IF local_bestIdx <> 0 THEN
                local_selected[local_bestIdx] := TRUE;
            END_IF;
        END_FOR;

        FOR local_i := 1 TO 5 DO
            pumpGroup[local_i].RunComd := local_selected[local_i];
        END_FOR;
    END_IF;
END_IF;

END_FUNCTION_BLOCK

(* ---- public-medium-01.raw_candidate_03.st ---- *)
(* ENGINEERING_CONTRACT
   - Mode FALSE=manual, TRUE=automatic (PUB001).
   - local_Running is retained run command: set by start OR previous running, cleared by stop; stop level wins (PUB002).
   - When local_Running=FALSE, all RunComd are FALSE (PUB002).
   - Manual running: each RunComd follows its current selection each scan (PUB001).
   - Automatic running: select 3 highest priority pumps, tie lower index; remaining stopped (PUB003).
   - priority/selection read-only; only RunComd written (PUB004).
*)
(* CONTRACT_RULES [] *)
TYPE ST_Pump :
STRUCT
    priority : INT;
    selection : BOOL;
    RunComd : BOOL;
END_STRUCT
END_TYPE;

FUNCTION_BLOCK FB_MultiPumpControl
VAR_INPUT
    mode : BOOL;
    start : BOOL;
    stop : BOOL;
END_VAR
VAR_IN_OUT
    pumpGroup : ARRAY[1..5] OF ST_Pump;
END_VAR
VAR
    local_Running : BOOL;
    local_selected : ARRAY[1..5] OF BOOL;
    local_bestIdx : INT;
    local_bestPrio : INT;
    local_i : INT;
    local_j : INT;
END_VAR

IF stop THEN
    local_Running := FALSE;
ELSE
    local_Running := local_Running OR start;
END_IF;

IF NOT local_Running THEN
    FOR local_i := 1 TO 5 DO
        pumpGroup[local_i].RunComd := FALSE;
    END_FOR;
ELSE
    IF NOT mode THEN
        FOR local_i := 1 TO 5 DO
            pumpGroup[local_i].RunComd := pumpGroup[local_i].selection;
        END_FOR;
    ELSE
        FOR local_i := 1 TO 5 DO
            local_selected[local_i] := FALSE;
        END_FOR;

        FOR local_j := 1 TO 3 DO
            local_bestIdx := 0;
            local_bestPrio := -32768;

            FOR local_i := 1 TO 5 DO
                IF NOT local_selected[local_i] THEN
                    IF (local_bestIdx = 0) OR (pumpGroup[local_i].priority > local_bestPrio) THEN
                        local_bestIdx := local_i;
                        local_bestPrio := pumpGroup[local_i].priority;
                    END_IF;
                END_IF;
            END_FOR;

            IF local_bestIdx <> 0 THEN
                local_selected[local_bestIdx] := TRUE;
            END_IF;
        END_FOR;

        FOR local_i := 1 TO 5 DO
            pumpGroup[local_i].RunComd := local_selected[local_i];
        END_FOR;
    END_IF;
END_IF;

END_FUNCTION_BLOCK

(* ---- public-medium-01.raw_candidate_04.st ---- *)
(* ENGINEERING_CONTRACT
   - Mode FALSE=manual, TRUE=automatic (PUB001).
   - Start is edge-triggered: a new FALSE->TRUE start pulse is required after stop release
     before pumps may run again; stop has priority over a level-held start (PUB001/PUB002).
   - local_Running is retained run state: set by rising edge of start while stop=FALSE,
     cleared immediately by stop=TRUE (PUB002).
   - When local_Running=FALSE, all RunComd are FALSE (PUB002).
   - Manual running: each RunComd follows its current selection each scan (PUB001).
   - Automatic running: select 3 highest priority pumps, tie lower index; remaining stopped (PUB003).
   - priority/selection read-only; only RunComd written (PUB004).
*)
(* CONTRACT_RULES [] *)
TYPE ST_Pump :
STRUCT
    priority : INT;
    selection : BOOL;
    RunComd : BOOL;
END_STRUCT
END_TYPE

FUNCTION_BLOCK FB_MultiPumpControl
VAR_INPUT
    mode : BOOL;
    start : BOOL;
    stop : BOOL;
END_VAR
VAR_IN_OUT
    pumpGroup : ARRAY[1..5] OF ST_Pump;
END_VAR
VAR
    local_Running : BOOL;
    local_selected : ARRAY[1..5] OF BOOL;
    local_bestIdx : INT;
    local_bestPrio : INT;
    local_i : INT;
    local_j : INT;
    local_rtStart : R_TRIG;
END_VAR

local_rtStart(CLK := start);

IF stop THEN
    local_Running := FALSE;
ELSE
    local_Running := local_Running OR local_rtStart.Q;
END_IF;

IF NOT local_Running THEN
    FOR local_i := 1 TO 5 DO
        pumpGroup[local_i].RunComd := FALSE;
    END_FOR;
ELSE
    IF NOT mode THEN
        FOR local_i := 1 TO 5 DO
            pumpGroup[local_i].RunComd := pumpGroup[local_i].selection;
        END_FOR;
    ELSE
        FOR local_i := 1 TO 5 DO
            local_selected[local_i] := FALSE;
        END_FOR;

        FOR local_j := 1 TO 3 DO
            local_bestIdx := 0;
            local_bestPrio := -32768;

            FOR local_i := 1 TO 5 DO
                IF NOT local_selected[local_i] THEN
                    IF (local_bestIdx = 0) OR (pumpGroup[local_i].priority > local_bestPrio) THEN
                        local_bestIdx := local_i;
                        local_bestPrio := pumpGroup[local_i].priority;
                    END_IF;
                END_IF;
            END_FOR;

            IF local_bestIdx <> 0 THEN
                local_selected[local_bestIdx] := TRUE;
            END_IF;
        END_FOR;

        FOR local_i := 1 TO 5 DO
            pumpGroup[local_i].RunComd := local_selected[local_i];
        END_FOR;
    END_IF;
END_IF;

END_FUNCTION_BLOCK

(* ---- public-medium-02.candidate_01.st ---- *)
TYPE ST_AnalogChannel :
STRUCT
    enable : BOOL;
    hiLIM : REAL;
    loLIM : REAL;
    bipolar : BOOL;
    measuringMode : INT;
    retVal : WORD;
    outputValue : REAL;
END_STRUCT
END_TYPE;

FUNCTION_BLOCK AnalogBatchProcessing
VAR_INPUT
    count : DINT;
END_VAR
VAR_INOUT
    analogValues : ARRAY[*] OF INT;
    channels : ARRAY[*] OF ST_AnalogChannel;
END_VAR
VAR
    tmp_i : DINT;
    tmp_process_count : DINT;
    tmp_analog_lower : DINT;
    tmp_channel_lower : DINT;
    tmp_analog_len : DINT;
    tmp_channel_len : DINT;
    tmp_raw : INT;
    tmp_raw_real : REAL;
    tmp_span : REAL;
    tmp_range : REAL;
END_VAR

(* ENGINEERING_CONTRACT
   Outputs:
   channels[].retVal : activation = enabled channel processed; retention = written only then; reset = none; priority = mode error before limit error; units: WORD.
   channels[].outputValue : activation = successful conversion only; retention = unchanged on skip/error/disabled; reset = none; units: REAL.
   Disabled channels: no writes.
   Mode 0 scaling boundaries: unipolar raw 0..27648 maps [loLIM,hiLIM], bipolar raw -27648..27648 maps [loLIM,hiLIM]; no clamping specified (PUB003).
   Mode 1/2 scale raw/10, raw/100 (PUB004, PUB005).
   Count represents ordinal positions from each array lower bound; caller valid 0..min lengths (PUB001). Cap invalid high count to available.
   Priority for invalid mode vs limit: invalid mode 16#8001 checked first, then limit 16#8002 (PUB006, PUB007).
*)

(* CONTRACT_RULES [] *)

tmp_analog_lower := LOWER_BOUND(analogValues, 1);
tmp_channel_lower := LOWER_BOUND(channels, 1);
tmp_analog_len := UPPER_BOUND(analogValues, 1) - tmp_analog_lower + 1;
tmp_channel_len := UPPER_BOUND(channels, 1) - tmp_channel_lower + 1;

IF count <= 0 THEN
    RETURN;
END_IF;

tmp_process_count := count;
IF tmp_process_count > tmp_analog_len THEN
    tmp_process_count := tmp_analog_len;
END_IF;
IF tmp_process_count > tmp_channel_len THEN
    tmp_process_count := tmp_channel_len;
END_IF;

FOR tmp_i := 0 TO tmp_process_count - 1 DO
    IF channels[tmp_channel_lower + tmp_i].enable THEN
        IF channels[tmp_channel_lower + tmp_i].measuringMode < 0 OR
           channels[tmp_channel_lower + tmp_i].measuringMode > 2 THEN
            channels[tmp_channel_lower + tmp_i].retVal := 16#8001;
        ELSIF channels[tmp_channel_lower + tmp_i].hiLIM <= channels[tmp_channel_lower + tmp_i].loLIM THEN
            channels[tmp_channel_lower + tmp_i].retVal := 16#8002;
        ELSE
            channels[tmp_channel_lower + tmp_i].retVal := 0;
            tmp_raw := analogValues[tmp_analog_lower + tmp_i];
            tmp_raw_real := TO_REAL(tmp_raw);
            CASE channels[tmp_channel_lower + tmp_i].measuringMode OF
                0:
                    tmp_span := channels[tmp_channel_lower + tmp_i].hiLIM - channels[tmp_channel_lower + tmp_i].loLIM;
                    IF channels[tmp_channel_lower + tmp_i].bipolar THEN
                        tmp_range := 55296.0;
                        channels[tmp_channel_lower + tmp_i].outputValue :=
                            channels[tmp_channel_lower + tmp_i].loLIM +
                            ((tmp_raw_real + 27648.0) / tmp_range) * tmp_span;
                    ELSE
                        tmp_range := 27648.0;
                        channels[tmp_channel_lower + tmp_i].outputValue :=
                            channels[tmp_channel_lower + tmp_i].loLIM +
                            (tmp_raw_real / tmp_range) * tmp_span;
                    END_IF;
                1:
                    channels[tmp_channel_lower + tmp_i].outputValue := tmp_raw_real / 10.0;
                2:
                    channels[tmp_channel_lower + tmp_i].outputValue := tmp_raw_real / 100.0;
            END_CASE;
        END_IF;
    END_IF;
END_FOR;

END_FUNCTION_BLOCK

(* ---- public-medium-02.candidate_02.st ---- *)
TYPE ST_AnalogChannel :
STRUCT
    enable : BOOL;
    hiLIM : REAL;
    loLIM : REAL;
    bipolar : BOOL;
    measuringMode : INT;
    retVal : WORD;
    outputValue : REAL;
END_STRUCT
END_TYPE;

FUNCTION_BLOCK AnalogBatchProcessing
VAR_INPUT
    count : DINT;
END_VAR
VAR_IN_OUT
    analogValues : ARRAY[*] OF INT;
    channels : ARRAY[*] OF ST_AnalogChannel;
END_VAR
VAR
    tmp_i : DINT;
    tmp_process_count : DINT;
    tmp_analog_lower : DINT;
    tmp_channel_lower : DINT;
    tmp_analog_len : DINT;
    tmp_channel_len : DINT;
    tmp_raw : INT;
    tmp_raw_real : REAL;
    tmp_span : REAL;
    tmp_range : REAL;
END_VAR

(* ENGINEERING_CONTRACT
   Outputs:
   channels[].retVal : activation = enabled channel processed; retention = written only then; reset = none; priority = mode error before limit error; units: WORD.
   channels[].outputValue : activation = successful conversion only; retention = unchanged on skip/error/disabled; reset = none; units: REAL.
   Disabled channels: no writes.
   Mode 0 scaling boundaries: unipolar raw 0..27648 maps [loLIM,hiLIM], bipolar raw -27648..27648 maps [loLIM,hiLIM]; no clamping specified (PUB003).
   Mode 1/2 scale raw/10, raw/100 (PUB004, PUB005).
   Count represents ordinal positions from each array lower bound; caller valid 0..min lengths (PUB001). Cap invalid high count to available.
   Priority for invalid mode vs limit: invalid mode 16#8001 checked first, then limit 16#8002 (PUB006, PUB007).
*)

(* CONTRACT_RULES [] *)

tmp_analog_lower := LOWER_BOUND(analogValues, 1);
tmp_channel_lower := LOWER_BOUND(channels, 1);
tmp_analog_len := UPPER_BOUND(analogValues, 1) - tmp_analog_lower + 1;
tmp_channel_len := UPPER_BOUND(channels, 1) - tmp_channel_lower + 1;

IF count <= 0 THEN
    RETURN;
END_IF;

tmp_process_count := count;
IF tmp_process_count > tmp_analog_len THEN
    tmp_process_count := tmp_analog_len;
END_IF;
IF tmp_process_count > tmp_channel_len THEN
    tmp_process_count := tmp_channel_len;
END_IF;

FOR tmp_i := 0 TO tmp_process_count - 1 DO
    IF channels[tmp_channel_lower + tmp_i].enable THEN
        IF channels[tmp_channel_lower + tmp_i].measuringMode < 0 OR
           channels[tmp_channel_lower + tmp_i].measuringMode > 2 THEN
            channels[tmp_channel_lower + tmp_i].retVal := 16#8001;
        ELSIF channels[tmp_channel_lower + tmp_i].hiLIM <= channels[tmp_channel_lower + tmp_i].loLIM THEN
            channels[tmp_channel_lower + tmp_i].retVal := 16#8002;
        ELSE
            channels[tmp_channel_lower + tmp_i].retVal := 0;
            tmp_raw := analogValues[tmp_analog_lower + tmp_i];
            tmp_raw_real := TO_REAL(tmp_raw);
            CASE channels[tmp_channel_lower + tmp_i].measuringMode OF
                0:
                    tmp_span := channels[tmp_channel_lower + tmp_i].hiLIM - channels[tmp_channel_lower + tmp_i].loLIM;
                    IF channels[tmp_channel_lower + tmp_i].bipolar THEN
                        tmp_range := 55296.0;
                        channels[tmp_channel_lower + tmp_i].outputValue :=
                            channels[tmp_channel_lower + tmp_i].loLIM +
                            ((tmp_raw_real + 27648.0) / tmp_range) * tmp_span;
                    ELSE
                        tmp_range := 27648.0;
                        channels[tmp_channel_lower + tmp_i].outputValue :=
                            channels[tmp_channel_lower + tmp_i].loLIM +
                            (tmp_raw_real / tmp_range) * tmp_span;
                    END_IF;
                1:
                    channels[tmp_channel_lower + tmp_i].outputValue := tmp_raw_real / 10.0;
                2:
                    channels[tmp_channel_lower + tmp_i].outputValue := tmp_raw_real / 100.0;
            END_CASE;
        END_IF;
    END_IF;
END_FOR;

END_FUNCTION_BLOCK
